Universal Robots URScript: FaiChun_9 Jan_6.script

def Machining1():
  # Default parameters:
  global speed_ms = 0.05
  global speed_rads = 0.75
  global accel_mss = 3
  global accel_radss = 1.2
  global blend_radius_m = 0.0003

  # Add subprograms here
  # Start of main program
  # Program generated by RoboDK v5.6.8 for UR10e on 10/01/2025 10:27:31
  # Using nominal kinematics.
  blend_radius_m = 0.0003
  speed_ms = 0.05
  # set_reference(p[0.325000, -0.070000, 0.000000, 0.000000, 0.000000, 0.000000])
  set_tcp(p[0.000000, 0.000000, 0.252000, 0.000000, 0.000000, 0.000000])
  # Show Tool
  movej([0.540600, -1.409576, -2.440611, -0.862202, 1.570796, 2.111396],accel_radss,speed_rads,0,blend_radius_m)
  movel([0.540600, -1.462244, -2.470081, -0.780064, 1.570796, 2.111396],accel_mss,speed_ms,0,blend_radius_m)
  #SetTool1
  #M_RunCode6
  #SetRPM60000
  speed_ms = 0.05
  #M_RunCode3
  movel([0.540600, -1.485155, -2.481004, -0.746230, 1.570796, 2.111396],accel_mss,speed_ms,0,blend_radius_m)
  speed_ms = 0.003
  movel([0.540600, -1.491068, -2.483663, -0.737658, 1.570796, 2.111396],accel_mss,speed_ms,0,blend_radius_m)
  speed_ms = 0.007
  movel([0.231188, -1.485347, -2.488632, -0.738410, 1.570796, 1.801984],accel_mss,speed_ms,0,blend_radius_m)
  movel([0.347864, -1.099241, -2.719319, -0.893829, 1.570796, 1.918660],accel_mss,speed_ms,0,blend_radius_m)
  movel([0.790744, -1.114546, -2.713470, -0.884373, 1.570796, 2.361541],accel_mss,speed_ms,0,blend_radius_m)
  movel([0.540600, -1.491068, -2.483663, -0.737658, 1.570796, 2.111396],accel_mss,speed_ms,0,blend_radius_m)
  speed_ms = 0.003
  movel([0.540600, -1.485155, -2.481004, -0.746230, 1.570796, 2.111396],accel_mss,speed_ms,0,blend_radius_m)
  speed_ms = 0.05
  movel([0.540600, -1.462244, -2.470081, -0.780064, 1.570796, 2.111396],accel_mss,speed_ms,0,blend_radius_m)
  #M_RunCode9
  movel([0.540492, -1.452284, -2.478323, -0.781782, 1.570796, 2.111289],accel_mss,speed_ms,0,blend_radius_m)
  #M_RunCode3
  movel([0.540492, -1.475406, -2.489363, -0.747620, 1.570796, 2.111289],accel_mss,speed_ms,0,blend_radius_m)
  speed_ms = 0.003
  movel([0.540492, -1.481377, -2.492050, -0.738962, 1.570796, 2.111289],accel_mss,speed_ms,0,blend_radius_m)
  speed_ms = 0.007
  movel([0.536155, -1.480632, -2.492689, -0.739069, 1.570796, 2.106951],accel_mss,speed_ms,0,blend_radius_m)
  movel([0.533586, -1.484990, -2.488940, -0.738459, 1.570796, 2.104382],accel_mss,speed_ms,0,blend_radius_m)
  movel([0.527159, -1.483935, -2.489850, -0.738604, 1.570796, 2.097955],accel_mss,speed_ms,0,blend_radius_m)
  movel([0.529703, -1.479563, -2.493604, -0.739223, 1.570796, 2.100499],accel_mss,speed_ms,0,blend_radius_m)
  movel([0.527435, -1.479199, -2.493915, -0.739276, 1.570796, 2.098231],accel_mss,speed_ms,0,blend_radius_m)
  movel([0.524898, -1.483575, -2.490161, -0.738654, 1.570796, 2.095694],accel_mss,speed_ms,0,blend_radius_m)
  movel([0.519478, -1.482738, -2.490881, -0.738770, 1.570796, 2.090274],accel_mss,speed_ms,0,blend_radius_m)
  movel([0.518427, -1.482577, -2.491019, -0.738793, 1.570796, 2.089223],accel_mss,speed_ms,0,blend_radius_m)
  movel([0.522154, -1.476073, -2.496578, -0.739738, 1.570796, 2.092951],accel_mss,speed_ms,0,blend_radius_m)
  movel([0.526552, -1.476753, -2.496000, -0.739636, 1.570796, 2.097348],accel_mss,speed_ms,0,blend_radius_m)
  movel([0.527881, -1.474461, -2.497945, -0.739983, 1.570796, 2.098677],accel_mss,speed_ms,0,blend_radius_m)
  movel([0.521180, -1.473430, -2.498818, -0.740141, 1.570796, 2.091976],accel_mss,speed_ms,0,blend_radius_m)
  movel([0.516149, -1.482240, -2.491309, -0.738840, 1.570796, 2.086946],accel_mss,speed_ms,0,blend_radius_m)
  movel([0.515092, -1.482086, -2.491441, -0.738862, 1.570796, 2.085888],accel_mss,speed_ms,0,blend_radius_m)
  movel([0.392568, -1.472171, -2.499881, -0.740337, 1.570796, 1.963364],accel_mss,speed_ms,0,blend_radius_m)
  movel([0.261942, -1.477589, -2.495288, -0.739512, 1.570796, 1.832738],accel_mss,speed_ms,0,blend_radius_m)
  movel([0.264591, -1.468670, -2.502825, -0.740895, 1.570796, 1.835387],accel_mss,speed_ms,0,blend_radius_m)
  movel([0.257067, -1.469444, -2.502175, -0.740770, 1.570796, 1.827863],accel_mss,speed_ms,0,blend_radius_m)
  movel([0.256391, -1.471766, -2.500222, -0.740401, 1.570796, 1.827188],accel_mss,speed_ms,0,blend_radius_m)
  movel([0.261332, -1.471251, -2.500656, -0.740482, 1.570796, 1.832129],accel_mss,speed_ms,0,blend_radius_m)
  movel([0.259390, -1.477836, -2.495078, -0.739475, 1.570796, 1.830187],accel_mss,speed_ms,0,blend_radius_m)
  movel([0.258210, -1.477956, -2.494975, -0.739458, 1.570796, 1.829007],accel_mss,speed_ms,0,blend_radius_m)
  movel([0.252127, -1.478591, -2.494434, -0.739364, 1.570796, 1.822923],accel_mss,speed_ms,0,blend_radius_m)
  movel([0.253398, -1.474162, -2.498199, -0.740029, 1.570796, 1.824194],accel_mss,speed_ms,0,blend_radius_m)
  movel([0.250836, -1.474438, -2.497965, -0.739986, 1.570796, 1.821633],accel_mss,speed_ms,0,blend_radius_m)
  movel([0.249578, -1.478866, -2.494199, -0.739324, 1.570796, 1.820375],accel_mss,speed_ms,0,blend_radius_m)
  movel([0.242307, -1.479680, -2.493504, -0.739206, 1.570796, 1.813103],accel_mss,speed_ms,0,blend_radius_m)
  movel([0.243527, -1.475262, -2.497266, -0.739861, 1.570796, 1.814323],accel_mss,speed_ms,0,blend_radius_m)
  movel([0.238589, -1.475844, -2.496772, -0.739773, 1.570796, 1.809385],accel_mss,speed_ms,0,blend_radius_m)
  movel([0.240380, -1.469260, -2.502330, -0.740799, 1.570796, 1.811176],accel_mss,speed_ms,0,blend_radius_m)
  movel([0.245358, -1.468668, -2.502826, -0.740895, 1.570796, 1.816154],accel_mss,speed_ms,0,blend_radius_m)
  movel([0.246004, -1.466343, -2.504771, -0.741276, 1.570796, 1.816800],accel_mss,speed_ms,0,blend_radius_m)
  movel([0.241015, -1.466936, -2.504276, -0.741178, 1.570796, 1.811811],accel_mss,speed_ms,0,blend_radius_m)
  movel([0.242546, -1.461356, -2.508913, -0.742121, 1.570796, 1.813342],accel_mss,speed_ms,0,blend_radius_m)
  movel([0.242845, -1.460267, -2.509812, -0.742310, 1.570796, 1.813642],accel_mss,speed_ms,0,blend_radius_m)
  movel([0.250292, -1.459376, -2.510546, -0.742467, 1.570796, 1.821088],accel_mss,speed_ms,0,blend_radius_m)
  movel([0.249014, -1.463897, -2.506806, -0.741685, 1.570796, 1.819810],accel_mss,speed_ms,0,blend_radius_m)
  movel([0.251610, -1.463600, -2.507053, -0.741736, 1.570796, 1.822406],accel_mss,speed_ms,0,blend_radius_m)
  movel([0.253577, -1.456716, -2.512732, -0.742941, 1.570796, 1.824373],accel_mss,speed_ms,0,blend_radius_m)
  movel([0.243495, -1.457910, -2.511752, -0.742727, 1.570796, 1.814291],accel_mss,speed_ms,0,blend_radius_m)
  movel([0.283133, -1.321596, -2.609965, -0.780829, 1.570796, 1.853929],accel_mss,speed_ms,0,blend_radius_m)
  movel([0.338490, -1.148112, -2.699863, -0.864413, 1.570796, 1.909286],accel_mss,speed_ms,0,blend_radius_m)
  movel([0.339093, -1.146307, -2.700623, -0.865459, 1.570796, 1.909889],accel_mss,speed_ms,0,blend_radius_m)
  movel([0.353258, -1.143604, -2.701755, -0.867030, 1.570796, 1.924055],accel_mss,speed_ms,0,blend_radius_m)
  movel([0.357266, -1.132009, -2.706527, -0.873852, 1.570796, 1.928063],accel_mss,speed_ms,0,blend_radius_m)
  movel([0.353555, -1.132710, -2.706243, -0.873436, 1.570796, 1.924351],accel_mss,speed_ms,0,blend_radius_m)
  movel([0.350931, -1.140355, -2.703106, -0.868929, 1.570796, 1.921727],accel_mss,speed_ms,0,blend_radius_m)
  movel([0.340411, -1.142384, -2.702263, -0.867742, 1.570796, 1.911208],accel_mss,speed_ms,0,blend_radius_m)
  movel([0.341015, -1.140566, -2.703018, -0.868805, 1.570796, 1.911811],accel_mss,speed_ms,0,blend_radius_m)
  movel([0.344182, -1.131093, -2.706899, -0.874397, 1.570796, 1.914978],accel_mss,speed_ms,0,blend_radius_m)
  movel([0.351373, -1.129671, -2.707474, -0.875244, 1.570796, 1.922170],accel_mss,speed_ms,0,blend_radius_m)
  movel([0.352747, -1.125647, -2.709091, -0.877652, 1.570796, 1.923543],accel_mss,speed_ms,0,blend_radius_m)
  movel([0.345526, -1.127083, -2.708515, -0.876791, 1.570796, 1.916323],accel_mss,speed_ms,0,blend_radius_m)
  movel([0.349422, -1.115504, -2.713097, -0.883789, 1.570796, 1.920218],accel_mss,speed_ms,0,blend_radius_m)
  movel([0.356727, -1.114025, -2.713673, -0.884691, 1.570796, 1.927524],accel_mss,speed_ms,0,blend_radius_m)
  movel([0.359466, -1.106053, -2.716742, -0.889593, 1.570796, 1.930262],accel_mss,speed_ms,0,blend_radius_m)
  movel([0.370357, -1.103908, -2.717558, -0.890922, 1.570796, 1.941153],accel_mss,speed_ms,0,blend_radius_m)
  movel([0.367527, -1.111926, -2.714487, -0.885976, 1.570796, 1.938324],accel_mss,speed_ms,0,blend_radius_m)
  movel([0.371310, -1.111216, -2.714761, -0.886412, 1.570796, 1.942106],accel_mss,speed_ms,0,blend_radius_m)
  movel([0.374169, -1.103183, -2.717833, -0.891372, 1.570796, 1.944966],accel_mss,speed_ms,0,blend_radius_m)
  movel([0.385027, -1.101192, -2.718585, -0.892612, 1.570796, 1.955823],accel_mss,speed_ms,0,blend_radius_m)
  movel([0.380684, -1.113104, -2.714031, -0.885255, 1.570796, 1.951481],accel_mss,speed_ms,0,blend_radius_m)
  movel([0.373438, -1.114398, -2.713528, -0.884463, 1.570796, 1.944234],accel_mss,speed_ms,0,blend_radius_m)
  movel([0.371969, -1.118508, -2.711920, -0.881961, 1.570796, 1.942765],accel_mss,speed_ms,0,blend_radius_m)
  movel([0.382929, -1.116581, -2.712676, -0.883132, 1.570796, 1.953725],accel_mss,speed_ms,0,blend_radius_m)
  movel([0.388829, -1.100520, -2.718838, -0.893030, 1.570796, 1.959625],accel_mss,speed_ms,0,blend_radius_m)
  movel([0.580174, -1.086020, -2.724199, -0.902169, 1.570796, 2.150970],accel_mss,speed_ms,0,blend_radius_m)
  movel([0.749145, -1.112705, -2.714185, -0.885499, 1.570796, 2.319942],accel_mss,speed_ms,0,blend_radius_m)
  movel([0.738673, -1.128310, -2.708023, -0.876057, 1.570796, 2.309469],accel_mss,speed_ms,0,blend_radius_m)
  movel([0.747236, -1.130824, -2.707008, -0.874557, 1.570796, 2.318032],accel_mss,speed_ms,0,blend_radius_m)
  movel([0.749941, -1.126842, -2.708612, -0.876935, 1.570796, 2.320738],accel_mss,speed_ms,0,blend_radius_m)
  movel([0.744304, -1.125159, -2.709286, -0.877945, 1.570796, 2.315100],accel_mss,speed_ms,0,blend_radius_m)
  movel([0.752109, -1.113600, -2.713838, -0.884951, 1.570796, 2.322905],accel_mss,speed_ms,0,blend_radius_m)
  movel([0.753475, -1.114012, -2.713678, -0.884699, 1.570796, 2.324272],accel_mss,speed_ms,0,blend_radius_m)
  movel([0.760489, -1.116181, -2.712832, -0.883375, 1.570796, 2.331285],accel_mss,speed_ms,0,blend_radius_m)
  movel([0.755172, -1.123962, -2.709763, -0.878664, 1.570796, 2.325968],accel_mss,speed_ms,0,blend_radius_m)
  movel([0.758077, -1.124873, -2.709400, -0.878116, 1.570796, 2.328873],accel_mss,speed_ms,0,blend_radius_m)
  movel([0.763409, -1.117111, -2.712468, -0.882809, 1.570796, 2.334206],accel_mss,speed_ms,0,blend_radius_m)
  movel([0.771667, -1.119832, -2.711399, -0.881158, 1.570796, 2.342463],accel_mss,speed_ms,0,blend_radius_m)
  movel([0.766309, -1.127539, -2.708332, -0.876518, 1.570796, 2.337105],accel_mss,speed_ms,0,blend_radius_m)
  movel([0.771815, -1.129393, -2.707586, -0.875410, 1.570796, 2.342612],accel_mss,speed_ms,0,blend_radius_m)
  movel([0.763990, -1.140583, -2.703011, -0.868795, 1.570796, 2.334786],accel_mss,speed_ms,0,blend_radius_m)
  movel([0.758513, -1.138781, -2.703756, -0.869852, 1.570796, 2.329309],accel_mss,speed_ms,0,blend_radius_m)
  movel([0.755817, -1.142675, -2.702142, -0.867572, 1.570796, 2.326613],accel_mss,speed_ms,0,blend_radius_m)
  movel([0.761284, -1.144460, -2.701397, -0.866532, 1.570796, 2.332081],accel_mss,speed_ms,0,blend_radius_m)
  movel([0.754898, -1.153625, -2.697523, -0.861241, 1.570796, 2.325695],accel_mss,speed_ms,0,blend_radius_m)
  movel([0.753674, -1.155384, -2.696769, -0.860235, 1.570796, 2.324470],accel_mss,speed_ms,0,blend_radius_m)
  movel([0.745605, -1.152827, -2.697863, -0.861698, 1.570796, 2.316402],accel_mss,speed_ms,0,blend_radius_m)
  movel([0.750697, -1.145425, -2.700993, -0.865971, 1.570796, 2.321494],accel_mss,speed_ms,0,blend_radius_m)
  movel([0.747837, -1.144533, -2.701367, -0.866489, 1.570796, 2.318634],accel_mss,speed_ms,0,blend_radius_m)
  movel([0.740145, -1.155770, -2.696604, -0.860015, 1.570796, 2.310941],accel_mss,speed_ms,0,blend_radius_m)
  movel([0.751042, -1.159170, -2.695138, -0.858082, 1.570796, 2.321838],accel_mss,speed_ms,0,blend_radius_m)
  movel([0.635581, -1.329799, -2.604798, -0.777792, 1.570796, 2.206378],accel_mss,speed_ms,0,blend_radius_m)
  movel([0.551105, -1.463690, -2.506978, -0.741720, 1.570796, 2.121901],accel_mss,speed_ms,0,blend_radius_m)
  movel([0.542267, -1.462159, -2.508248, -0.741982, 1.570796, 2.113063],accel_mss,speed_ms,0,blend_radius_m)
  movel([0.538244, -1.468952, -2.502588, -0.740849, 1.570796, 2.109040],accel_mss,speed_ms,0,blend_radius_m)
  movel([0.540528, -1.469337, -2.502265, -0.740787, 1.570796, 2.111324],accel_mss,speed_ms,0,blend_radius_m)
  movel([0.543178, -1.464878, -2.505991, -0.741520, 1.570796, 2.113974],accel_mss,speed_ms,0,blend_radius_m)
  movel([0.549694, -1.466015, -2.505044, -0.741330, 1.570796, 2.120491],accel_mss,speed_ms,0,blend_radius_m)
  movel([0.549048, -1.467088, -2.504148, -0.741153, 1.570796, 2.119844],accel_mss,speed_ms,0,blend_radius_m)
  movel([0.545741, -1.472593, -2.499525, -0.740271, 1.570796, 2.116537],accel_mss,speed_ms,0,blend_radius_m)
  movel([0.541370, -1.471831, -2.500168, -0.740390, 1.570796, 2.112167],accel_mss,speed_ms,0,blend_radius_m)
  movel([0.540008, -1.474125, -2.498230, -0.740034, 1.570796, 2.110804],accel_mss,speed_ms,0,blend_radius_m)
  movel([0.544370, -1.474884, -2.497587, -0.739918, 1.570796, 2.115167],accel_mss,speed_ms,0,blend_radius_m)
  movel([0.540492, -1.481377, -2.492050, -0.738962, 1.570796, 2.111289],accel_mss,speed_ms,0,blend_radius_m)
  speed_ms = 0.003
  movel([0.540492, -1.475406, -2.489363, -0.747620, 1.570796, 2.111289],accel_mss,speed_ms,0,blend_radius_m)
  speed_ms = 0.05
  movel([0.540492, -1.452284, -2.478323, -0.781782, 1.570796, 2.111289],accel_mss,speed_ms,0,blend_radius_m)
  #M_RunCode9
  movel([0.384099, -1.143946, -2.667631, -0.900812, 1.570796, 1.954895],accel_mss,speed_ms,0,blend_radius_m)
  #M_RunCode3
  movel([0.384099, -1.171719, -2.682638, -0.858032, 1.570796, 1.954895],accel_mss,speed_ms,0,blend_radius_m)
  speed_ms = 0.003
  movel([0.384099, -1.179045, -2.686328, -0.847016, 1.570796, 1.954895],accel_mss,speed_ms,0,blend_radius_m)
  speed_ms = 0.007
  movel([0.371180, -1.190123, -2.681237, -0.841029, 1.570796, 1.941977],accel_mss,speed_ms,0,blend_radius_m)
  movel([0.353670, -1.164627, -2.692759, -0.855002, 1.570796, 1.924466],accel_mss,speed_ms,0,blend_radius_m)
  movel([0.354978, -1.163450, -2.693275, -0.855664, 1.570796, 1.925774],accel_mss,speed_ms,0,blend_radius_m)
  movel([0.358519, -1.160754, -2.694450, -0.857185, 1.570796, 1.929315],accel_mss,speed_ms,0,blend_radius_m)
  movel([0.362422, -1.158698, -2.695342, -0.858349, 1.570796, 1.933218],accel_mss,speed_ms,0,blend_radius_m)
  movel([0.366466, -1.157207, -2.695985, -0.859196, 1.570796, 1.937262],accel_mss,speed_ms,0,blend_radius_m)
  movel([0.370429, -1.156192, -2.696422, -0.859774, 1.570796, 1.941225],accel_mss,speed_ms,0,blend_radius_m)
  movel([0.380760, -1.154569, -2.697119, -0.860701, 1.570796, 1.951557],accel_mss,speed_ms,0,blend_radius_m)
  movel([0.390288, -1.153250, -2.697683, -0.861456, 1.570796, 1.961084],accel_mss,speed_ms,0,blend_radius_m)
  movel([0.393974, -1.152407, -2.698042, -0.861939, 1.570796, 1.964770],accel_mss,speed_ms,0,blend_radius_m)
  movel([0.397663, -1.151161, -2.698572, -0.862655, 1.570796, 1.968460],accel_mss,speed_ms,0,blend_radius_m)
  movel([0.401177, -1.149434, -2.699305, -0.863650, 1.570796, 1.971974],accel_mss,speed_ms,0,blend_radius_m)
  movel([0.404336, -1.147153, -2.700267, -0.864968, 1.570796, 1.975133],accel_mss,speed_ms,0,blend_radius_m)
  movel([0.407651, -1.143740, -2.701698, -0.866951, 1.570796, 1.978447],accel_mss,speed_ms,0,blend_radius_m)
  movel([0.408788, -1.142051, -2.702402, -0.867936, 1.570796, 1.979584],accel_mss,speed_ms,0,blend_radius_m)
  movel([0.409576, -1.140378, -2.703096, -0.868915, 1.570796, 1.980372],accel_mss,speed_ms,0,blend_radius_m)
  movel([0.410196, -1.137359, -2.704342, -0.870688, 1.570796, 1.980993],accel_mss,speed_ms,0,blend_radius_m)
  movel([0.409610, -1.134976, -2.705319, -0.872094, 1.570796, 1.980407],accel_mss,speed_ms,0,blend_radius_m)
  movel([0.408647, -1.133848, -2.705779, -0.872762, 1.570796, 1.979444],accel_mss,speed_ms,0,blend_radius_m)
  movel([0.407469, -1.133422, -2.705953, -0.873014, 1.570796, 1.978266],accel_mss,speed_ms,0,blend_radius_m)
  movel([0.406201, -1.133623, -2.705871, -0.872895, 1.570796, 1.976997],accel_mss,speed_ms,0,blend_radius_m)
  movel([0.404968, -1.134393, -2.705557, -0.872439, 1.570796, 1.975765],accel_mss,speed_ms,0,blend_radius_m)
  movel([0.403605, -1.136287, -2.704782, -0.871320, 1.570796, 1.974401],accel_mss,speed_ms,0,blend_radius_m)
  movel([0.402385, -1.138186, -2.704001, -0.870202, 1.570796, 1.973181],accel_mss,speed_ms,0,blend_radius_m)
  movel([0.400444, -1.140181, -2.703178, -0.869031, 1.570796, 1.971241],accel_mss,speed_ms,0,blend_radius_m)
  movel([0.397817, -1.141968, -2.702436, -0.867985, 1.570796, 1.968613],accel_mss,speed_ms,0,blend_radius_m)
  movel([0.395422, -1.142572, -2.702185, -0.867632, 1.570796, 1.966218],accel_mss,speed_ms,0,blend_radius_m)
  movel([0.393436, -1.142139, -2.702365, -0.867885, 1.570796, 1.964232],accel_mss,speed_ms,0,blend_radius_m)
  movel([0.392041, -1.140812, -2.702916, -0.868661, 1.570796, 1.962837],accel_mss,speed_ms,0,blend_radius_m)
  movel([0.391392, -1.138828, -2.703737, -0.869824, 1.570796, 1.962188],accel_mss,speed_ms,0,blend_radius_m)
  movel([0.391640, -1.136425, -2.704725, -0.871238, 1.570796, 1.962436],accel_mss,speed_ms,0,blend_radius_m)
  movel([0.392852, -1.133853, -2.705777, -0.872758, 1.570796, 1.963649],accel_mss,speed_ms,0,blend_radius_m)
  movel([0.395102, -1.131371, -2.706786, -0.874232, 1.570796, 1.965898],accel_mss,speed_ms,0,blend_radius_m)
  movel([0.397379, -1.129656, -2.707480, -0.875253, 1.570796, 1.968175],accel_mss,speed_ms,0,blend_radius_m)
  movel([0.399624, -1.128553, -2.707925, -0.875911, 1.570796, 1.970420],accel_mss,speed_ms,0,blend_radius_m)
  movel([0.401834, -1.128068, -2.708120, -0.876202, 1.570796, 1.972630],accel_mss,speed_ms,0,blend_radius_m)
  movel([0.404002, -1.128203, -2.708066, -0.876121, 1.570796, 1.974798],accel_mss,speed_ms,0,blend_radius_m)
  movel([0.406053, -1.128886, -2.707791, -0.875713, 1.570796, 1.976850],accel_mss,speed_ms,0,blend_radius_m)
  movel([0.407900, -1.130046, -2.707322, -0.875020, 1.570796, 1.978697],accel_mss,speed_ms,0,blend_radius_m)
  movel([0.410999, -1.133777, -2.705808, -0.872804, 1.570796, 1.981795],accel_mss,speed_ms,0,blend_radius_m)
  movel([0.412374, -1.136716, -2.704606, -0.871067, 1.570796, 1.983170],accel_mss,speed_ms,0,blend_radius_m)
  movel([0.413232, -1.139861, -2.703310, -0.869218, 1.570796, 1.984028],accel_mss,speed_ms,0,blend_radius_m)
  movel([0.413580, -1.143201, -2.701923, -0.867265, 1.570796, 1.984376],accel_mss,speed_ms,0,blend_radius_m)
  movel([0.413422, -1.146734, -2.700444, -0.865211, 1.570796, 1.984218],accel_mss,speed_ms,0,blend_radius_m)
  movel([0.412572, -1.150319, -2.698930, -0.863140, 1.570796, 1.983368],accel_mss,speed_ms,0,blend_radius_m)
  movel([0.410842, -1.153822, -2.697438, -0.861128, 1.570796, 1.981638],accel_mss,speed_ms,0,blend_radius_m)
  movel([0.408237, -1.157248, -2.695968, -0.859173, 1.570796, 1.979033],accel_mss,speed_ms,0,blend_radius_m)
  movel([0.404766, -1.160594, -2.694520, -0.857275, 1.570796, 1.975563],accel_mss,speed_ms,0,blend_radius_m)
  movel([0.401302, -1.163173, -2.693396, -0.855820, 1.570796, 1.972098],accel_mss,speed_ms,0,blend_radius_m)
  movel([0.397796, -1.165070, -2.692565, -0.854754, 1.570796, 1.968592],accel_mss,speed_ms,0,blend_radius_m)
  movel([0.394330, -1.166408, -2.691977, -0.854005, 1.570796, 1.965126],accel_mss,speed_ms,0,blend_radius_m)
  movel([0.391000, -1.167299, -2.691584, -0.853506, 1.570796, 1.961796],accel_mss,speed_ms,0,blend_radius_m)
  movel([0.383085, -1.168489, -2.691058, -0.852842, 1.570796, 1.953882],accel_mss,speed_ms,0,blend_radius_m)
  movel([0.375587, -1.169704, -2.690520, -0.852166, 1.570796, 1.946383],accel_mss,speed_ms,0,blend_radius_m)
  movel([0.372556, -1.170542, -2.690147, -0.851700, 1.570796, 1.943353],accel_mss,speed_ms,0,blend_radius_m)
  movel([0.369459, -1.171768, -2.689601, -0.851020, 1.570796, 1.940255],accel_mss,speed_ms,0,blend_radius_m)
  movel([0.366399, -1.173459, -2.688845, -0.850085, 1.570796, 1.937196],accel_mss,speed_ms,0,blend_radius_m)
  movel([0.363487, -1.175689, -2.687844, -0.848856, 1.570796, 1.934283],accel_mss,speed_ms,0,blend_radius_m)
  movel([0.364141, -1.176646, -2.687413, -0.848330, 1.570796, 1.934937],accel_mss,speed_ms,0,blend_radius_m)
  movel([0.366146, -1.179126, -2.686291, -0.846972, 1.570796, 1.936943],accel_mss,speed_ms,0,blend_radius_m)
  movel([0.368319, -1.180933, -2.685469, -0.845986, 1.570796, 1.939115],accel_mss,speed_ms,0,blend_radius_m)
  movel([0.370657, -1.182078, -2.684947, -0.845364, 1.570796, 1.941454],accel_mss,speed_ms,0,blend_radius_m)
  movel([0.373172, -1.182554, -2.684729, -0.845105, 1.570796, 1.943968],accel_mss,speed_ms,0,blend_radius_m)
  movel([0.375804, -1.182447, -2.684778, -0.845164, 1.570796, 1.946600],accel_mss,speed_ms,0,blend_radius_m)
  movel([0.378498, -1.181829, -2.685061, -0.845499, 1.570796, 1.949294],accel_mss,speed_ms,0,blend_radius_m)
  movel([0.381261, -1.180696, -2.685577, -0.846115, 1.570796, 1.952058],accel_mss,speed_ms,0,blend_radius_m)
  movel([0.384099, -1.179045, -2.686328, -0.847016, 1.570796, 1.954895],accel_mss,speed_ms,0,blend_radius_m)
  speed_ms = 0.003
  movel([0.384099, -1.171719, -2.682638, -0.858032, 1.570796, 1.954895],accel_mss,speed_ms,0,blend_radius_m)
  speed_ms = 0.05
  movel([0.384099, -1.143946, -2.667631, -0.900812, 1.570796, 1.954895],accel_mss,speed_ms,0,blend_radius_m)
  #M_RunCode9
  movel([0.391981, -1.155983, -2.662339, -0.894068, 1.570796, 1.962777],accel_mss,speed_ms,0,blend_radius_m)
  #M_RunCode3
  movel([0.391981, -1.183682, -2.677188, -0.851519, 1.570796, 1.962777],accel_mss,speed_ms,0,blend_radius_m)
  speed_ms = 0.003
  movel([0.391981, -1.190981, -2.680837, -0.840571, 1.570796, 1.962777],accel_mss,speed_ms,0,blend_radius_m)
  speed_ms = 0.007
  movel([0.401981, -1.182312, -2.684840, -0.845237, 1.570796, 1.972777],accel_mss,speed_ms,0,blend_radius_m)
  movel([0.412364, -1.173981, -2.688611, -0.849796, 1.570796, 1.983160],accel_mss,speed_ms,0,blend_radius_m)
  movel([0.420048, -1.168557, -2.691028, -0.852804, 1.570796, 1.990844],accel_mss,speed_ms,0,blend_radius_m)
  movel([0.422893, -1.166993, -2.691719, -0.853677, 1.570796, 1.993689],accel_mss,speed_ms,0,blend_radius_m)
  movel([0.425127, -1.166238, -2.692052, -0.854100, 1.570796, 1.995924],accel_mss,speed_ms,0,blend_radius_m)
  movel([0.426748, -1.166298, -2.692025, -0.854066, 1.570796, 1.997544],accel_mss,speed_ms,0,blend_radius_m)
  movel([0.427747, -1.167174, -2.691639, -0.853576, 1.570796, 1.998543],accel_mss,speed_ms,0,blend_radius_m)
  movel([0.428014, -1.168646, -2.690988, -0.852754, 1.570796, 1.998811],accel_mss,speed_ms,0,blend_radius_m)
  movel([0.427442, -1.170502, -2.690165, -0.851722, 1.570796, 1.998239],accel_mss,speed_ms,0,blend_radius_m)
  movel([0.426031, -1.172734, -2.689170, -0.850485, 1.570796, 1.996828],accel_mss,speed_ms,0,blend_radius_m)
  movel([0.423792, -1.175342, -2.688001, -0.849047, 1.570796, 1.994589],accel_mss,speed_ms,0,blend_radius_m)
  movel([0.416876, -1.181935, -2.685012, -0.845442, 1.570796, 1.987672],accel_mss,speed_ms,0,blend_radius_m)
  movel([0.406811, -1.190510, -2.681057, -0.840823, 1.570796, 1.977607],accel_mss,speed_ms,0,blend_radius_m)
  movel([0.396637, -1.198599, -2.677252, -0.836537, 1.570796, 1.967434],accel_mss,speed_ms,0,blend_radius_m)
  movel([0.389261, -1.203802, -2.674767, -0.833820, 1.570796, 1.960057],accel_mss,speed_ms,0,blend_radius_m)
  movel([0.386540, -1.205311, -2.674041, -0.833037, 1.570796, 1.957337],accel_mss,speed_ms,0,blend_radius_m)
  movel([0.384392, -1.206055, -2.673682, -0.832652, 1.570796, 1.955188],accel_mss,speed_ms,0,blend_radius_m)
  movel([0.382806, -1.206040, -2.673689, -0.832660, 1.570796, 1.953602],accel_mss,speed_ms,0,blend_radius_m)
  movel([0.381784, -1.205259, -2.674066, -0.833064, 1.570796, 1.952580],accel_mss,speed_ms,0,blend_radius_m)
  movel([0.381444, -1.203906, -2.674717, -0.833765, 1.570796, 1.952240],accel_mss,speed_ms,0,blend_radius_m)
  movel([0.381917, -1.202164, -2.675553, -0.834672, 1.570796, 1.952713],accel_mss,speed_ms,0,blend_radius_m)
  movel([0.383201, -1.200030, -2.676572, -0.835787, 1.570796, 1.953998],accel_mss,speed_ms,0,blend_radius_m)
  movel([0.385310, -1.197499, -2.677774, -0.837116, 1.570796, 1.956107],accel_mss,speed_ms,0,blend_radius_m)
  movel([0.391981, -1.190981, -2.680837, -0.840571, 1.570796, 1.962777],accel_mss,speed_ms,0,blend_radius_m)
  speed_ms = 0.003
  movel([0.391981, -1.183682, -2.677188, -0.851519, 1.570796, 1.962777],accel_mss,speed_ms,0,blend_radius_m)
  speed_ms = 0.05
  movel([0.391981, -1.155983, -2.662339, -0.894068, 1.570796, 1.962777],accel_mss,speed_ms,0,blend_radius_m)
  #M_RunCode9
  movel([0.382534, -1.154364, -2.663059, -0.894966, 1.570796, 1.953331],accel_mss,speed_ms,0,blend_radius_m)
  #M_RunCode3
  movel([0.382534, -1.182074, -2.677929, -0.852386, 1.570796, 1.953331],accel_mss,speed_ms,0,blend_radius_m)
  speed_ms = 0.003
  movel([0.382534, -1.189377, -2.681584, -0.841428, 1.570796, 1.953331],accel_mss,speed_ms,0,blend_radius_m)
  speed_ms = 0.007
  movel([0.384510, -1.186300, -2.683009, -0.843080, 1.570796, 1.955306],accel_mss,speed_ms,0,blend_radius_m)
  movel([0.386914, -1.183128, -2.684467, -0.844794, 1.570796, 1.957710],accel_mss,speed_ms,0,blend_radius_m)
  movel([0.389736, -1.179922, -2.685929, -0.846537, 1.570796, 1.960532],accel_mss,speed_ms,0,blend_radius_m)
  movel([0.392976, -1.176687, -2.687394, -0.848307, 1.570796, 1.963773],accel_mss,speed_ms,0,blend_radius_m)
  movel([0.396639, -1.173419, -2.688863, -0.850106, 1.570796, 1.967435],accel_mss,speed_ms,0,blend_radius_m)
  movel([0.400453, -1.170358, -2.690229, -0.851802, 1.570796, 1.971250],accel_mss,speed_ms,0,blend_radius_m)
  movel([0.404137, -1.167738, -2.691390, -0.853261, 1.570796, 1.974933],accel_mss,speed_ms,0,blend_radius_m)
  movel([0.407690, -1.165566, -2.692347, -0.854476, 1.570796, 1.978486],accel_mss,speed_ms,0,blend_radius_m)
  movel([0.411102, -1.163850, -2.693100, -0.855439, 1.570796, 1.981898],accel_mss,speed_ms,0,blend_radius_m)
  movel([0.414313, -1.162590, -2.693651, -0.856149, 1.570796, 1.985110],accel_mss,speed_ms,0,blend_radius_m)
  movel([0.417262, -1.161790, -2.694000, -0.856600, 1.570796, 1.988058],accel_mss,speed_ms,0,blend_radius_m)
  movel([0.419951, -1.161449, -2.694148, -0.856792, 1.570796, 1.990747],accel_mss,speed_ms,0,blend_radius_m)
  movel([0.422369, -1.161571, -2.694095, -0.856723, 1.570796, 1.993165],accel_mss,speed_ms,0,blend_radius_m)
  movel([0.424501, -1.162118, -2.693856, -0.856414, 1.570796, 1.995297],accel_mss,speed_ms,0,blend_radius_m)
  movel([0.426315, -1.163065, -2.693443, -0.855881, 1.570796, 1.997111],accel_mss,speed_ms,0,blend_radius_m)
  movel([0.427820, -1.164408, -2.692856, -0.855126, 1.570796, 1.998617],accel_mss,speed_ms,0,blend_radius_m)
  movel([0.429009, -1.166139, -2.692095, -0.854155, 1.570796, 1.999805],accel_mss,speed_ms,0,blend_radius_m)
  movel([0.429838, -1.168160, -2.691203, -0.853025, 1.570796, 2.000634],accel_mss,speed_ms,0,blend_radius_m)
  movel([0.430255, -1.170379, -2.690220, -0.851791, 1.570796, 2.001051],accel_mss,speed_ms,0,blend_radius_m)
  movel([0.430265, -1.172781, -2.689149, -0.850459, 1.570796, 2.001061],accel_mss,speed_ms,0,blend_radius_m)
  movel([0.429867, -1.175374, -2.687986, -0.849029, 1.570796, 2.000663],accel_mss,speed_ms,0,blend_radius_m)
  movel([0.429057, -1.178111, -2.686751, -0.847527, 1.570796, 1.999853],accel_mss,speed_ms,0,blend_radius_m)
  movel([0.427818, -1.180961, -2.685457, -0.845972, 1.570796, 1.998614],accel_mss,speed_ms,0,blend_radius_m)
  movel([0.426158, -1.183915, -2.684106, -0.844368, 1.570796, 1.996955],accel_mss,speed_ms,0,blend_radius_m)
  movel([0.424077, -1.186979, -2.682695, -0.842715, 1.570796, 1.994873],accel_mss,speed_ms,0,blend_radius_m)
  movel([0.421597, -1.190091, -2.681252, -0.841046, 1.570796, 1.992393],accel_mss,speed_ms,0,blend_radius_m)
  movel([0.418745, -1.193188, -2.679805, -0.839396, 1.570796, 1.989541],accel_mss,speed_ms,0,blend_radius_m)
  movel([0.415518, -1.196270, -2.678355, -0.837764, 1.570796, 1.986314],accel_mss,speed_ms,0,blend_radius_m)
  movel([0.411919, -1.199346, -2.676897, -0.836146, 1.570796, 1.982715],accel_mss,speed_ms,0,blend_radius_m)
  movel([0.408214, -1.202196, -2.675537, -0.834655, 1.570796, 1.979010],accel_mss,speed_ms,0,blend_radius_m)
  movel([0.404666, -1.204615, -2.674377, -0.833398, 1.570796, 1.975463],accel_mss,speed_ms,0,blend_radius_m)
  movel([0.401273, -1.206606, -2.673416, -0.832367, 1.570796, 1.972069],accel_mss,speed_ms,0,blend_radius_m)
  movel([0.398024, -1.208172, -2.672657, -0.831560, 1.570796, 1.968821],accel_mss,speed_ms,0,blend_radius_m)
  movel([0.394967, -1.209327, -2.672096, -0.830966, 1.570796, 1.965763],accel_mss,speed_ms,0,blend_radius_m)
  movel([0.392151, -1.210070, -2.671734, -0.830585, 1.570796, 1.962947],accel_mss,speed_ms,0,blend_radius_m)
  movel([0.389569, -1.210403, -2.671572, -0.830414, 1.570796, 1.960365],accel_mss,speed_ms,0,blend_radius_m)
  movel([0.387217, -1.210331, -2.671607, -0.830451, 1.570796, 1.958013],accel_mss,speed_ms,0,blend_radius_m)
  movel([0.385124, -1.209875, -2.671829, -0.830685, 1.570796, 1.955920],accel_mss,speed_ms,0,blend_radius_m)
  movel([0.383309, -1.209055, -2.672228, -0.831106, 1.570796, 1.954105],accel_mss,speed_ms,0,blend_radius_m)
  movel([0.381774, -1.207869, -2.672804, -0.831715, 1.570796, 1.952571],accel_mss,speed_ms,0,blend_radius_m)
  movel([0.380519, -1.206319, -2.673555, -0.832516, 1.570796, 1.951316],accel_mss,speed_ms,0,blend_radius_m)
  movel([0.379600, -1.204481, -2.674441, -0.833467, 1.570796, 1.950397],accel_mss,speed_ms,0,blend_radius_m)
  movel([0.379072, -1.202440, -2.675421, -0.834528, 1.570796, 1.949868],accel_mss,speed_ms,0,blend_radius_m)
  movel([0.378939, -1.200190, -2.676496, -0.835703, 1.570796, 1.949735],accel_mss,speed_ms,0,blend_radius_m)
  movel([0.379206, -1.197729, -2.677665, -0.836995, 1.570796, 1.950002],accel_mss,speed_ms,0,blend_radius_m)
  movel([0.379886, -1.195089, -2.678912, -0.838388, 1.570796, 1.950682],accel_mss,speed_ms,0,blend_radius_m)
  movel([0.380993, -1.192308, -2.680217, -0.839864, 1.570796, 1.951790],accel_mss,speed_ms,0,blend_radius_m)
  movel([0.382534, -1.189377, -2.681584, -0.841428, 1.570796, 1.953331],accel_mss,speed_ms,0,blend_radius_m)
  speed_ms = 0.003
  movel([0.382534, -1.182074, -2.677929, -0.852386, 1.570796, 1.953331],accel_mss,speed_ms,0,blend_radius_m)
  speed_ms = 0.05
  movel([0.382534, -1.154364, -2.663059, -0.894966, 1.570796, 1.953331],accel_mss,speed_ms,0,blend_radius_m)
  #M_RunCode9
  movel([0.494383, -1.389930, -2.526626, -0.795833, 1.570796, 2.065179],accel_mss,speed_ms,0,blend_radius_m)
  #M_RunCode3
  movel([0.494383, -1.414326, -2.538424, -0.759639, 1.570796, 2.065179],accel_mss,speed_ms,0,blend_radius_m)
  speed_ms = 0.003
  movel([0.494383, -1.420647, -2.541300, -0.750441, 1.570796, 2.065179],accel_mss,speed_ms,0,blend_radius_m)
  speed_ms = 0.007
  movel([0.497081, -1.419373, -2.542274, -0.750742, 1.570796, 2.067877],accel_mss,speed_ms,0,blend_radius_m)
  movel([0.499941, -1.418639, -2.542833, -0.750917, 1.570796, 2.070737],accel_mss,speed_ms,0,blend_radius_m)
  movel([0.502829, -1.418338, -2.543062, -0.750988, 1.570796, 2.073625],accel_mss,speed_ms,0,blend_radius_m)
  movel([0.505605, -1.418366, -2.543041, -0.750982, 1.570796, 2.076401],accel_mss,speed_ms,0,blend_radius_m)
  movel([0.512719, -1.419167, -2.542431, -0.750791, 1.570796, 2.083515],accel_mss,speed_ms,0,blend_radius_m)
  movel([0.519252, -1.420019, -2.541780, -0.750589, 1.570796, 2.090049],accel_mss,speed_ms,0,blend_radius_m)
  movel([0.521814, -1.420108, -2.541713, -0.750569, 1.570796, 2.092610],accel_mss,speed_ms,0,blend_radius_m)
  movel([0.524418, -1.419908, -2.541865, -0.750616, 1.570796, 2.095214],accel_mss,speed_ms,0,blend_radius_m)
  movel([0.526952, -1.419333, -2.542304, -0.750752, 1.570796, 2.097748],accel_mss,speed_ms,0,blend_radius_m)
  movel([0.529302, -1.418300, -2.543092, -0.750998, 1.570796, 2.100099],accel_mss,speed_ms,0,blend_radius_m)
  movel([0.531866, -1.416496, -2.544463, -0.751431, 1.570796, 2.102662],accel_mss,speed_ms,0,blend_radius_m)
  movel([0.532796, -1.415514, -2.545207, -0.751668, 1.570796, 2.103592],accel_mss,speed_ms,0,blend_radius_m)
  movel([0.533494, -1.414477, -2.545991, -0.751921, 1.570796, 2.104290],accel_mss,speed_ms,0,blend_radius_m)
  movel([0.534215, -1.412459, -2.547513, -0.752417, 1.570796, 2.105012],accel_mss,speed_ms,0,blend_radius_m)
  movel([0.534067, -1.410667, -2.548859, -0.752863, 1.570796, 2.104864],accel_mss,speed_ms,0,blend_radius_m)
  movel([0.533541, -1.409690, -2.549591, -0.753108, 1.570796, 2.104338],accel_mss,speed_ms,0,blend_radius_m)
  movel([0.532799, -1.409167, -2.549982, -0.753240, 1.570796, 2.103596],accel_mss,speed_ms,0,blend_radius_m)
  movel([0.531934, -1.409071, -2.550054, -0.753264, 1.570796, 2.102730],accel_mss,speed_ms,0,blend_radius_m)
  movel([0.531038, -1.409381, -2.549822, -0.753186, 1.570796, 2.101834],accel_mss,speed_ms,0,blend_radius_m)
  movel([0.529935, -1.410463, -2.549012, -0.752914, 1.570796, 2.100731],accel_mss,speed_ms,0,blend_radius_m)
  movel([0.528924, -1.411578, -2.548175, -0.752636, 1.570796, 2.099720],accel_mss,speed_ms,0,blend_radius_m)
  movel([0.527424, -1.412624, -2.547389, -0.752376, 1.570796, 2.098220],accel_mss,speed_ms,0,blend_radius_m)
  movel([0.525483, -1.413399, -2.546805, -0.752185, 1.570796, 2.096280],accel_mss,speed_ms,0,blend_radius_m)
  movel([0.523822, -1.413373, -2.546824, -0.752192, 1.570796, 2.094618],accel_mss,speed_ms,0,blend_radius_m)
  movel([0.522542, -1.412689, -2.547340, -0.752360, 1.570796, 2.093338],accel_mss,speed_ms,0,blend_radius_m)
  movel([0.521753, -1.411480, -2.548249, -0.752660, 1.570796, 2.092549],accel_mss,speed_ms,0,blend_radius_m)
  movel([0.521531, -1.409947, -2.549399, -0.753043, 1.570796, 2.092327],accel_mss,speed_ms,0,blend_radius_m)
  movel([0.521953, -1.408286, -2.550640, -0.753462, 1.570796, 2.092749],accel_mss,speed_ms,0,blend_radius_m)
  movel([0.523034, -1.406692, -2.551828, -0.753868, 1.570796, 2.093830],accel_mss,speed_ms,0,blend_radius_m)
  movel([0.524792, -1.405362, -2.552817, -0.754210, 1.570796, 2.095589],accel_mss,speed_ms,0,blend_radius_m)
  movel([0.526486, -1.404585, -2.553393, -0.754411, 1.570796, 2.097282],accel_mss,speed_ms,0,blend_radius_m)
  movel([0.528091, -1.404236, -2.553652, -0.754502, 1.570796, 2.098888],accel_mss,speed_ms,0,blend_radius_m)
  movel([0.529608, -1.404316, -2.553592, -0.754481, 1.570796, 2.100405],accel_mss,speed_ms,0,blend_radius_m)
  movel([0.531035, -1.404826, -2.553214, -0.754349, 1.570796, 2.101831],accel_mss,speed_ms,0,blend_radius_m)
  movel([0.532324, -1.405698, -2.552567, -0.754124, 1.570796, 2.103120],accel_mss,speed_ms,0,blend_radius_m)
  movel([0.533433, -1.406868, -2.551698, -0.753824, 1.570796, 2.104229],accel_mss,speed_ms,0,blend_radius_m)
  movel([0.535111, -1.410082, -2.549298, -0.753010, 1.570796, 2.105907],accel_mss,speed_ms,0,blend_radius_m)
  movel([0.535730, -1.412414, -2.547547, -0.752428, 1.570796, 2.106526],accel_mss,speed_ms,0,blend_radius_m)
  movel([0.535987, -1.414790, -2.545754, -0.751845, 1.570796, 2.106783],accel_mss,speed_ms,0,blend_radius_m)
  movel([0.535884, -1.417214, -2.543918, -0.751258, 1.570796, 2.106680],accel_mss,speed_ms,0,blend_radius_m)
  movel([0.535424, -1.419683, -2.542037, -0.750669, 1.570796, 2.106221],accel_mss,speed_ms,0,blend_radius_m)
  movel([0.534495, -1.422065, -2.540215, -0.750110, 1.570796, 2.105292],accel_mss,speed_ms,0,blend_radius_m)
  movel([0.532980, -1.424234, -2.538547, -0.749607, 1.570796, 2.103776],accel_mss,speed_ms,0,blend_radius_m)
  movel([0.530887, -1.426191, -2.537037, -0.749161, 1.570796, 2.101683],accel_mss,speed_ms,0,blend_radius_m)
  movel([0.528209, -1.427943, -2.535681, -0.748765, 1.570796, 2.099005],accel_mss,speed_ms,0,blend_radius_m)
  movel([0.525614, -1.429150, -2.534743, -0.748496, 1.570796, 2.096411],accel_mss,speed_ms,0,blend_radius_m)
  movel([0.523054, -1.429866, -2.534186, -0.748337, 1.570796, 2.093850],accel_mss,speed_ms,0,blend_radius_m)
  movel([0.520575, -1.430192, -2.533932, -0.748265, 1.570796, 2.091372],accel_mss,speed_ms,0,blend_radius_m)
  movel([0.518236, -1.430218, -2.533912, -0.748259, 1.570796, 2.089032],accel_mss,speed_ms,0,blend_radius_m)
  movel([0.512764, -1.429613, -2.534383, -0.748393, 1.570796, 2.083560],accel_mss,speed_ms,0,blend_radius_m)
  movel([0.507570, -1.429093, -2.534787, -0.748508, 1.570796, 2.078366],accel_mss,speed_ms,0,blend_radius_m)
  movel([0.505430, -1.429133, -2.534757, -0.748500, 1.570796, 2.076226],accel_mss,speed_ms,0,blend_radius_m)
  movel([0.503200, -1.429440, -2.534518, -0.748432, 1.570796, 2.073996],accel_mss,speed_ms,0,blend_radius_m)
  movel([0.500938, -1.430091, -2.534011, -0.748287, 1.570796, 2.071735],accel_mss,speed_ms,0,blend_radius_m)
  movel([0.498716, -1.431164, -2.533174, -0.748051, 1.570796, 2.069512],accel_mss,speed_ms,0,blend_radius_m)
  movel([0.499050, -1.431983, -2.532534, -0.747872, 1.570796, 2.069846],accel_mss,speed_ms,0,blend_radius_m)
  movel([0.500128, -1.434162, -2.530827, -0.747400, 1.570796, 2.070924],accel_mss,speed_ms,0,blend_radius_m)
  movel([0.501395, -1.435883, -2.529473, -0.747032, 1.570796, 2.072191],accel_mss,speed_ms,0,blend_radius_m)
  movel([0.502857, -1.437147, -2.528476, -0.746765, 1.570796, 2.073653],accel_mss,speed_ms,0,blend_radius_m)
  movel([0.504510, -1.437959, -2.527835, -0.746595, 1.570796, 2.075306],accel_mss,speed_ms,0,blend_radius_m)
  movel([0.506311, -1.438363, -2.527515, -0.746511, 1.570796, 2.077107],accel_mss,speed_ms,0,blend_radius_m)
  movel([0.508208, -1.438409, -2.527479, -0.746501, 1.570796, 2.079004],accel_mss,speed_ms,0,blend_radius_m)
  movel([0.510207, -1.438094, -2.527728, -0.746567, 1.570796, 2.081003],accel_mss,speed_ms,0,blend_radius_m)
  movel([0.512309, -1.437419, -2.528261, -0.746708, 1.570796, 2.083106],accel_mss,speed_ms,0,blend_radius_m)
  movel([0.502315, -1.443102, -2.523747, -0.745540, 1.570796, 2.073111],accel_mss,speed_ms,0,blend_radius_m)
  movel([0.493365, -1.421248, -2.540841, -0.750300, 1.570796, 2.064162],accel_mss,speed_ms,0,blend_radius_m)
  movel([0.494383, -1.420647, -2.541300, -0.750441, 1.570796, 2.065179],accel_mss,speed_ms,0,blend_radius_m)
  speed_ms = 0.003
  movel([0.494383, -1.414326, -2.538424, -0.759639, 1.570796, 2.065179],accel_mss,speed_ms,0,blend_radius_m)
  speed_ms = 0.05
  movel([0.494383, -1.389930, -2.526626, -0.795833, 1.570796, 2.065179],accel_mss,speed_ms,0,blend_radius_m)
  #M_RunCode9
  movel([0.509612, -1.412120, -2.510078, -0.790191, 1.570796, 2.080409],accel_mss,speed_ms,0,blend_radius_m)
  #M_RunCode3
  movel([0.509612, -1.436073, -2.521602, -0.754714, 1.570796, 2.080409],accel_mss,speed_ms,0,blend_radius_m)
  speed_ms = 0.003
  movel([0.509612, -1.442272, -2.524410, -0.745707, 1.570796, 2.080409],accel_mss,speed_ms,0,blend_radius_m)
  speed_ms = 0.007
  movel([0.511490, -1.441522, -2.525007, -0.745860, 1.570796, 2.082287],accel_mss,speed_ms,0,blend_radius_m)
  movel([0.513128, -1.441532, -2.525000, -0.745858, 1.570796, 2.083924],accel_mss,speed_ms,0,blend_radius_m)
  movel([0.514398, -1.442178, -2.524485, -0.745726, 1.570796, 2.085195],accel_mss,speed_ms,0,blend_radius_m)
  movel([0.515181, -1.443333, -2.523562, -0.745493, 1.570796, 2.085977],accel_mss,speed_ms,0,blend_radius_m)
  movel([0.515399, -1.444801, -2.522388, -0.745200, 1.570796, 2.086195],accel_mss,speed_ms,0,blend_radius_m)
  movel([0.514982, -1.446386, -2.521116, -0.744887, 1.570796, 2.085779],accel_mss,speed_ms,0,blend_radius_m)
  movel([0.513938, -1.447896, -2.519900, -0.744592, 1.570796, 2.084734],accel_mss,speed_ms,0,blend_radius_m)
  movel([0.512272, -1.449136, -2.518900, -0.744353, 1.570796, 2.083068],accel_mss,speed_ms,0,blend_radius_m)
  movel([0.510726, -1.449811, -2.518354, -0.744224, 1.570796, 2.081522],accel_mss,speed_ms,0,blend_radius_m)
  movel([0.509449, -1.450009, -2.518194, -0.744186, 1.570796, 2.080246],accel_mss,speed_ms,0,blend_radius_m)
  movel([0.508135, -1.450311, -2.517949, -0.744128, 1.570796, 2.078931],accel_mss,speed_ms,0,blend_radius_m)
  movel([0.507400, -1.450916, -2.517460, -0.744014, 1.570796, 2.078197],accel_mss,speed_ms,0,blend_radius_m)
  movel([0.506930, -1.451756, -2.516778, -0.743855, 1.570796, 2.077727],accel_mss,speed_ms,0,blend_radius_m)
  movel([0.506762, -1.452683, -2.516025, -0.743681, 1.570796, 2.077558],accel_mss,speed_ms,0,blend_radius_m)
  movel([0.506927, -1.453558, -2.515312, -0.743519, 1.570796, 2.077723],accel_mss,speed_ms,0,blend_radius_m)
  movel([0.507485, -1.454522, -2.514526, -0.743341, 1.570796, 2.078282],accel_mss,speed_ms,0,blend_radius_m)
  movel([0.508303, -1.455228, -2.513950, -0.743211, 1.570796, 2.079099],accel_mss,speed_ms,0,blend_radius_m)
  movel([0.509379, -1.455675, -2.513584, -0.743130, 1.570796, 2.080176],accel_mss,speed_ms,0,blend_radius_m)
  movel([0.510712, -1.455870, -2.513425, -0.743094, 1.570796, 2.081508],accel_mss,speed_ms,0,blend_radius_m)
  movel([0.512224, -1.455797, -2.513485, -0.743108, 1.570796, 2.083021],accel_mss,speed_ms,0,blend_radius_m)
  movel([0.513839, -1.455450, -2.513768, -0.743171, 1.570796, 2.084635],accel_mss,speed_ms,0,blend_radius_m)
  movel([0.515560, -1.454826, -2.514278, -0.743285, 1.570796, 2.086356],accel_mss,speed_ms,0,blend_radius_m)
  movel([0.517386, -1.453926, -2.515013, -0.743451, 1.570796, 2.088182],accel_mss,speed_ms,0,blend_radius_m)
  movel([0.520257, -1.451945, -2.516624, -0.743819, 1.570796, 2.091053],accel_mss,speed_ms,0,blend_radius_m)
  movel([0.522585, -1.449475, -2.518626, -0.744288, 1.570796, 2.093382],accel_mss,speed_ms,0,blend_radius_m)
  movel([0.523520, -1.448065, -2.519765, -0.744560, 1.570796, 2.094316],accel_mss,speed_ms,0,blend_radius_m)
  movel([0.524260, -1.446552, -2.520982, -0.744854, 1.570796, 2.095056],accel_mss,speed_ms,0,blend_radius_m)
  movel([0.525158, -1.443210, -2.523661, -0.745518, 1.570796, 2.095955],accel_mss,speed_ms,0,blend_radius_m)
  movel([0.525179, -1.439539, -2.526583, -0.746267, 1.570796, 2.095975],accel_mss,speed_ms,0,blend_radius_m)
  movel([0.524211, -1.435637, -2.529668, -0.747085, 1.570796, 2.095007],accel_mss,speed_ms,0,blend_radius_m)
  movel([0.539789, -1.427052, -2.536371, -0.748966, 1.570796, 2.110585],accel_mss,speed_ms,0,blend_radius_m)
  movel([0.545461, -1.443958, -2.523063, -0.745368, 1.570796, 2.116257],accel_mss,speed_ms,0,blend_radius_m)
  movel([0.535452, -1.449327, -2.518746, -0.744316, 1.570796, 2.106249],accel_mss,speed_ms,0,blend_radius_m)
  movel([0.537620, -1.447411, -2.520291, -0.744687, 1.570796, 2.108416],accel_mss,speed_ms,0,blend_radius_m)
  movel([0.539396, -1.445076, -2.522167, -0.745145, 1.570796, 2.110192],accel_mss,speed_ms,0,blend_radius_m)
  movel([0.540687, -1.442436, -2.524279, -0.745674, 1.570796, 2.111484],accel_mss,speed_ms,0,blend_radius_m)
  movel([0.541406, -1.439606, -2.526530, -0.746253, 1.570796, 2.112203],accel_mss,speed_ms,0,blend_radius_m)
  movel([0.541489, -1.436695, -2.528833, -0.746861, 1.570796, 2.112285],accel_mss,speed_ms,0,blend_radius_m)
  movel([0.540874, -1.433817, -2.531098, -0.747474, 1.570796, 2.111670],accel_mss,speed_ms,0,blend_radius_m)
  movel([0.529435, -1.440058, -2.526171, -0.746160, 1.570796, 2.100232],accel_mss,speed_ms,0,blend_radius_m)
  movel([0.530293, -1.443522, -2.523411, -0.745455, 1.570796, 2.101089],accel_mss,speed_ms,0,blend_radius_m)
  movel([0.530471, -1.447177, -2.520480, -0.744732, 1.570796, 2.101268],accel_mss,speed_ms,0,blend_radius_m)
  movel([0.529866, -1.450823, -2.517535, -0.744031, 1.570796, 2.100662],accel_mss,speed_ms,0,blend_radius_m)
  movel([0.529229, -1.452573, -2.516114, -0.743702, 1.570796, 2.100025],accel_mss,speed_ms,0,blend_radius_m)
  movel([0.528372, -1.454274, -2.514729, -0.743386, 1.570796, 2.099168],accel_mss,speed_ms,0,blend_radius_m)
  movel([0.527276, -1.455875, -2.513420, -0.743093, 1.570796, 2.098072],accel_mss,speed_ms,0,blend_radius_m)
  movel([0.525923, -1.457328, -2.512230, -0.742831, 1.570796, 2.096719],accel_mss,speed_ms,0,blend_radius_m)
  movel([0.524317, -1.458631, -2.511159, -0.742598, 1.570796, 2.095113],accel_mss,speed_ms,0,blend_radius_m)
  movel([0.522454, -1.459792, -2.510204, -0.742393, 1.570796, 2.093250],accel_mss,speed_ms,0,blend_radius_m)
  movel([0.520506, -1.460724, -2.509434, -0.742230, 1.570796, 2.091302],accel_mss,speed_ms,0,blend_radius_m)
  movel([0.518643, -1.461347, -2.508920, -0.742122, 1.570796, 2.089440],accel_mss,speed_ms,0,blend_radius_m)
  movel([0.516862, -1.461661, -2.508660, -0.742068, 1.570796, 2.087658],accel_mss,speed_ms,0,blend_radius_m)
  movel([0.515163, -1.461668, -2.508654, -0.742067, 1.570796, 2.085960],accel_mss,speed_ms,0,blend_radius_m)
  movel([0.512100, -1.460952, -2.509246, -0.742191, 1.570796, 2.082897],accel_mss,speed_ms,0,blend_radius_m)
  movel([0.509548, -1.459390, -2.510535, -0.742464, 1.570796, 2.080345],accel_mss,speed_ms,0,blend_radius_m)
  movel([0.507542, -1.457189, -2.512344, -0.742856, 1.570796, 2.078338],accel_mss,speed_ms,0,blend_radius_m)
  movel([0.506120, -1.454557, -2.514498, -0.743334, 1.570796, 2.076917],accel_mss,speed_ms,0,blend_radius_m)
  movel([0.505558, -1.452516, -2.516160, -0.743713, 1.570796, 2.076354],accel_mss,speed_ms,0,blend_radius_m)
  movel([0.505383, -1.450221, -2.518022, -0.744145, 1.570796, 2.076179],accel_mss,speed_ms,0,blend_radius_m)
  movel([0.505659, -1.447865, -2.519926, -0.744598, 1.570796, 2.076455],accel_mss,speed_ms,0,blend_radius_m)
  movel([0.506446, -1.445637, -2.521718, -0.745034, 1.570796, 2.077243],accel_mss,speed_ms,0,blend_radius_m)
  movel([0.507761, -1.443713, -2.523259, -0.745417, 1.570796, 2.078557],accel_mss,speed_ms,0,blend_radius_m)
  movel([0.509612, -1.442272, -2.524410, -0.745707, 1.570796, 2.080409],accel_mss,speed_ms,0,blend_radius_m)
  speed_ms = 0.003
  movel([0.509612, -1.436073, -2.521602, -0.754714, 1.570796, 2.080409],accel_mss,speed_ms,0,blend_radius_m)
  speed_ms = 0.05
  movel([0.509612, -1.412120, -2.510078, -0.790191, 1.570796, 2.080409],accel_mss,speed_ms,0,blend_radius_m)
  #M_RunCode9
  movel([0.517025, -1.320922, -2.573739, -0.817728, 1.570796, 2.087821],accel_mss,speed_ms,0,blend_radius_m)
  #M_RunCode3
  movel([0.517025, -1.346591, -2.586414, -0.779384, 1.570796, 2.087821],accel_mss,speed_ms,0,blend_radius_m)
  speed_ms = 0.003
  movel([0.517025, -1.353271, -2.589511, -0.769607, 1.570796, 2.087821],accel_mss,speed_ms,0,blend_radius_m)
  speed_ms = 0.007
  movel([0.513857, -1.353859, -2.589119, -0.769412, 1.570796, 2.084654],accel_mss,speed_ms,0,blend_radius_m)
  movel([0.510784, -1.353806, -2.589154, -0.769429, 1.570796, 2.081580],accel_mss,speed_ms,0,blend_radius_m)
  movel([0.507871, -1.353220, -2.589545, -0.769624, 1.570796, 2.078668],accel_mss,speed_ms,0,blend_radius_m)
  movel([0.505181, -1.352209, -2.590219, -0.769961, 1.570796, 2.075978],accel_mss,speed_ms,0,blend_radius_m)
  movel([0.502784, -1.350876, -2.591105, -0.770407, 1.570796, 2.073580],accel_mss,speed_ms,0,blend_radius_m)
  movel([0.504597, -1.347224, -2.593522, -0.771643, 1.570796, 2.075394],accel_mss,speed_ms,0,blend_radius_m)
  movel([0.507463, -1.343318, -2.596086, -0.772985, 1.570796, 2.078259],accel_mss,speed_ms,0,blend_radius_m)
  movel([0.511084, -1.339508, -2.598566, -0.774315, 1.570796, 2.081881],accel_mss,speed_ms,0,blend_radius_m)
  movel([0.515153, -1.336160, -2.600729, -0.775499, 1.570796, 2.085949],accel_mss,speed_ms,0,blend_radius_m)
  movel([0.519346, -1.333645, -2.602345, -0.776399, 1.570796, 2.090142],accel_mss,speed_ms,0,blend_radius_m)
  movel([0.521387, -1.332816, -2.602876, -0.776698, 1.570796, 2.092183],accel_mss,speed_ms,0,blend_radius_m)
  movel([0.523335, -1.332335, -2.603183, -0.776871, 1.570796, 2.094131],accel_mss,speed_ms,0,blend_radius_m)
  movel([0.525151, -1.332246, -2.603239, -0.776903, 1.570796, 2.095947],accel_mss,speed_ms,0,blend_radius_m)
  movel([0.526785, -1.332598, -2.603015, -0.776776, 1.570796, 2.097581],accel_mss,speed_ms,0,blend_radius_m)
  movel([0.528204, -1.333429, -2.602483, -0.776477, 1.570796, 2.099000],accel_mss,speed_ms,0,blend_radius_m)
  movel([0.529362, -1.334787, -2.601613, -0.775989, 1.570796, 2.100158],accel_mss,speed_ms,0,blend_radius_m)
  movel([0.530223, -1.337369, -2.599950, -0.775070, 1.570796, 2.101019],accel_mss,speed_ms,0,blend_radius_m)
  movel([0.529939, -1.340263, -2.598076, -0.774050, 1.570796, 2.100735],accel_mss,speed_ms,0,blend_radius_m)
  movel([0.528649, -1.343348, -2.596066, -0.772975, 1.570796, 2.099445],accel_mss,speed_ms,0,blend_radius_m)
  movel([0.526489, -1.346505, -2.593995, -0.771889, 1.570796, 2.097286],accel_mss,speed_ms,0,blend_radius_m)
  movel([0.523400, -1.349714, -2.591876, -0.770799, 1.570796, 2.094196],accel_mss,speed_ms,0,blend_radius_m)
  movel([0.520226, -1.351927, -2.590407, -0.770055, 1.570796, 2.091022],accel_mss,speed_ms,0,blend_radius_m)
  movel([0.517025, -1.353271, -2.589511, -0.769607, 1.570796, 2.087821],accel_mss,speed_ms,0,blend_radius_m)
  speed_ms = 0.003
  movel([0.517025, -1.346591, -2.586414, -0.779384, 1.570796, 2.087821],accel_mss,speed_ms,0,blend_radius_m)
  speed_ms = 0.05
  movel([0.517025, -1.320922, -2.573739, -0.817728, 1.570796, 2.087821],accel_mss,speed_ms,0,blend_radius_m)
  #M_RunCode9
  movel([0.612042, -1.222485, -2.630373, -0.859530, 1.570796, 2.182838],accel_mss,speed_ms,0,blend_radius_m)
  #M_RunCode3
  movel([0.612042, -1.249578, -2.644343, -0.818468, 1.570796, 2.182838],accel_mss,speed_ms,0,blend_radius_m)
  speed_ms = 0.003
  movel([0.612042, -1.256679, -2.647767, -0.807942, 1.570796, 2.182838],accel_mss,speed_ms,0,blend_radius_m)
  speed_ms = 0.007
  movel([0.610850, -1.255352, -2.648485, -0.808552, 1.570796, 2.181646],accel_mss,speed_ms,0,blend_radius_m)
  movel([0.610180, -1.253548, -2.649458, -0.809383, 1.570796, 2.180977],accel_mss,speed_ms,0,blend_radius_m)
  movel([0.609813, -1.251505, -2.650554, -0.810330, 1.570796, 2.180609],accel_mss,speed_ms,0,blend_radius_m)
  movel([0.610746, -1.251259, -2.650686, -0.810444, 1.570796, 2.181542],accel_mss,speed_ms,0,blend_radius_m)
  movel([0.611268, -1.251665, -2.650468, -0.810256, 1.570796, 2.182064],accel_mss,speed_ms,0,blend_radius_m)
  movel([0.611926, -1.252076, -2.650248, -0.810065, 1.570796, 2.182722],accel_mss,speed_ms,0,blend_radius_m)
  movel([0.613261, -1.251850, -2.650369, -0.810170, 1.570796, 2.184057],accel_mss,speed_ms,0,blend_radius_m)
  movel([0.614772, -1.251013, -2.650818, -0.810559, 1.570796, 2.185568],accel_mss,speed_ms,0,blend_radius_m)
  movel([0.616233, -1.249908, -2.651408, -0.811073, 1.570796, 2.187029],accel_mss,speed_ms,0,blend_radius_m)
  movel([0.618237, -1.248311, -2.652258, -0.811820, 1.570796, 2.189033],accel_mss,speed_ms,0,blend_radius_m)
  movel([0.617947, -1.245637, -2.653675, -0.813076, 1.570796, 2.188743],accel_mss,speed_ms,0,blend_radius_m)
  movel([0.616923, -1.243875, -2.654605, -0.813909, 1.570796, 2.187719],accel_mss,speed_ms,0,blend_radius_m)
  movel([0.616065, -1.243468, -2.654819, -0.814102, 1.570796, 2.186862],accel_mss,speed_ms,0,blend_radius_m)
  movel([0.614938, -1.243449, -2.654829, -0.814111, 1.570796, 2.185734],accel_mss,speed_ms,0,blend_radius_m)
  movel([0.613515, -1.243869, -2.654608, -0.813912, 1.570796, 2.184311],accel_mss,speed_ms,0,blend_radius_m)
  movel([0.611773, -1.244776, -2.654130, -0.813483, 1.570796, 2.182570],accel_mss,speed_ms,0,blend_radius_m)
  movel([0.612499, -1.242950, -2.655091, -0.814348, 1.570796, 2.183296],accel_mss,speed_ms,0,blend_radius_m)
  movel([0.613329, -1.241381, -2.655914, -0.815094, 1.570796, 2.184125],accel_mss,speed_ms,0,blend_radius_m)
  movel([0.613825, -1.240829, -2.656203, -0.815357, 1.570796, 2.184622],accel_mss,speed_ms,0,blend_radius_m)
  movel([0.614394, -1.240506, -2.656371, -0.815511, 1.570796, 2.185191],accel_mss,speed_ms,0,blend_radius_m)
  movel([0.615825, -1.240771, -2.656233, -0.815385, 1.570796, 2.186622],accel_mss,speed_ms,0,blend_radius_m)
  movel([0.617921, -1.242529, -2.655312, -0.814548, 1.570796, 2.188718],accel_mss,speed_ms,0,blend_radius_m)
  movel([0.619316, -1.245004, -2.654010, -0.813375, 1.570796, 2.190112],accel_mss,speed_ms,0,blend_radius_m)
  movel([0.619584, -1.246454, -2.653244, -0.812692, 1.570796, 2.190380],accel_mss,speed_ms,0,blend_radius_m)
  movel([0.619474, -1.248016, -2.652415, -0.811958, 1.570796, 2.190270],accel_mss,speed_ms,0,blend_radius_m)
  movel([0.618929, -1.249665, -2.651537, -0.811187, 1.570796, 2.189725],accel_mss,speed_ms,0,blend_radius_m)
  movel([0.617880, -1.251383, -2.650619, -0.810386, 1.570796, 2.188676],accel_mss,speed_ms,0,blend_radius_m)
  movel([0.616504, -1.250348, -2.651173, -0.810868, 1.570796, 2.187301],accel_mss,speed_ms,0,blend_radius_m)
  movel([0.613987, -1.257295, -2.647433, -0.807660, 1.570796, 2.184783],accel_mss,speed_ms,0,blend_radius_m)
  movel([0.612042, -1.256679, -2.647767, -0.807942, 1.570796, 2.182838],accel_mss,speed_ms,0,blend_radius_m)
  speed_ms = 0.003
  movel([0.612042, -1.249578, -2.644343, -0.818468, 1.570796, 2.182838],accel_mss,speed_ms,0,blend_radius_m)
  speed_ms = 0.05
  movel([0.612042, -1.222485, -2.630373, -0.859530, 1.570796, 2.182838],accel_mss,speed_ms,0,blend_radius_m)
  #M_RunCode9
  movel([0.591456, -1.174119, -2.654087, -0.884183, 1.570796, 2.162252],accel_mss,speed_ms,0,blend_radius_m)
  #M_RunCode3
  movel([0.591456, -1.201686, -2.668697, -0.842006, 1.570796, 2.162252],accel_mss,speed_ms,0,blend_radius_m)
  speed_ms = 0.003
  movel([0.591456, -1.208939, -2.672285, -0.831165, 1.570796, 2.162252],accel_mss,speed_ms,0,blend_radius_m)
  speed_ms = 0.007
  movel([0.588359, -1.211205, -2.671180, -0.830004, 1.570796, 2.159155],accel_mss,speed_ms,0,blend_radius_m)
  movel([0.585138, -1.213198, -2.670204, -0.828987, 1.570796, 2.155934],accel_mss,speed_ms,0,blend_radius_m)
  movel([0.581822, -1.214884, -2.669375, -0.828130, 1.570796, 2.152618],accel_mss,speed_ms,0,blend_radius_m)
  movel([0.578445, -1.216225, -2.668713, -0.827451, 1.570796, 2.149242],accel_mss,speed_ms,0,blend_radius_m)
  movel([0.575048, -1.217185, -2.668237, -0.826966, 1.570796, 2.145844],accel_mss,speed_ms,0,blend_radius_m)
  movel([0.573345, -1.217319, -2.668171, -0.826899, 1.570796, 2.144141],accel_mss,speed_ms,0,blend_radius_m)
  movel([0.571660, -1.217172, -2.668244, -0.826973, 1.570796, 2.142456],accel_mss,speed_ms,0,blend_radius_m)
  movel([0.570140, -1.217053, -2.668303, -0.827033, 1.570796, 2.140936],accel_mss,speed_ms,0,blend_radius_m)
  movel([0.568941, -1.217262, -2.668200, -0.826928, 1.570796, 2.139737],accel_mss,speed_ms,0,blend_radius_m)
  movel([0.566873, -1.218693, -2.667489, -0.826207, 1.570796, 2.137669],accel_mss,speed_ms,0,blend_radius_m)
  movel([0.564147, -1.221009, -2.666335, -0.825045, 1.570796, 2.134944],accel_mss,speed_ms,0,blend_radius_m)
  movel([0.561318, -1.223454, -2.665109, -0.823826, 1.570796, 2.132115],accel_mss,speed_ms,0,blend_radius_m)
  movel([0.558932, -1.225284, -2.664188, -0.822917, 1.570796, 2.129728],accel_mss,speed_ms,0,blend_radius_m)
  movel([0.554225, -1.227961, -2.662833, -0.821596, 1.570796, 2.125021],accel_mss,speed_ms,0,blend_radius_m)
  movel([0.550026, -1.229677, -2.661959, -0.820752, 1.570796, 2.120823],accel_mss,speed_ms,0,blend_radius_m)
  movel([0.546288, -1.230531, -2.661524, -0.820334, 1.570796, 2.117084],accel_mss,speed_ms,0,blend_radius_m)
  movel([0.542964, -1.230613, -2.661482, -0.820294, 1.570796, 2.113760],accel_mss,speed_ms,0,blend_radius_m)
  movel([0.540020, -1.230006, -2.661792, -0.820591, 1.570796, 2.110816],accel_mss,speed_ms,0,blend_radius_m)
  movel([0.537407, -1.228804, -2.662404, -0.821181, 1.570796, 2.108203],accel_mss,speed_ms,0,blend_radius_m)
  movel([0.535098, -1.227083, -2.663278, -0.822028, 1.570796, 2.105894],accel_mss,speed_ms,0,blend_radius_m)
  movel([0.533056, -1.224929, -2.664367, -0.823093, 1.570796, 2.103852],accel_mss,speed_ms,0,blend_radius_m)
  movel([0.529627, -1.219666, -2.667005, -0.825718, 1.570796, 2.100423],accel_mss,speed_ms,0,blend_radius_m)
  movel([0.526861, -1.213687, -2.669964, -0.828738, 1.570796, 2.097657],accel_mss,speed_ms,0,blend_radius_m)
  movel([0.522289, -1.202428, -2.675427, -0.834534, 1.570796, 2.093085],accel_mss,speed_ms,0,blend_radius_m)
  movel([0.519671, -1.197902, -2.677583, -0.836904, 1.570796, 2.090467],accel_mss,speed_ms,0,blend_radius_m)
  movel([0.516029, -1.193158, -2.679819, -0.839412, 1.570796, 2.086825],accel_mss,speed_ms,0,blend_radius_m)
  movel([0.511507, -1.188478, -2.682001, -0.841910, 1.570796, 2.082304],accel_mss,speed_ms,0,blend_radius_m)
  movel([0.506261, -1.184167, -2.683990, -0.844232, 1.570796, 2.077057],accel_mss,speed_ms,0,blend_radius_m)
  movel([0.500453, -1.180515, -2.685660, -0.846214, 1.570796, 2.071249],accel_mss,speed_ms,0,blend_radius_m)
  movel([0.494265, -1.177818, -2.686884, -0.847687, 1.570796, 2.065061],accel_mss,speed_ms,0,blend_radius_m)
  movel([0.487893, -1.176356, -2.687544, -0.848489, 1.570796, 2.058690],accel_mss,speed_ms,0,blend_radius_m)
  movel([0.484702, -1.176171, -2.687627, -0.848591, 1.570796, 2.055498],accel_mss,speed_ms,0,blend_radius_m)
  movel([0.481544, -1.176394, -2.687527, -0.848468, 1.570796, 2.052340],accel_mss,speed_ms,0,blend_radius_m)
  movel([0.478145, -1.177057, -2.687228, -0.848105, 1.570796, 2.048941],accel_mss,speed_ms,0,blend_radius_m)
  movel([0.474068, -1.178233, -2.686696, -0.847460, 1.570796, 2.044865],accel_mss,speed_ms,0,blend_radius_m)
  movel([0.469550, -1.179944, -2.685919, -0.846525, 1.570796, 2.040347],accel_mss,speed_ms,0,blend_radius_m)
  movel([0.464822, -1.182215, -2.684884, -0.845290, 1.570796, 2.035619],accel_mss,speed_ms,0,blend_radius_m)
  movel([0.460129, -1.185051, -2.683584, -0.843754, 1.570796, 2.030925],accel_mss,speed_ms,0,blend_radius_m)
  movel([0.455702, -1.188467, -2.682006, -0.841916, 1.570796, 2.026499],accel_mss,speed_ms,0,blend_radius_m)
  movel([0.451783, -1.192465, -2.680144, -0.839780, 1.570796, 2.022579],accel_mss,speed_ms,0,blend_radius_m)
  movel([0.450084, -1.194681, -2.679104, -0.838604, 1.570796, 2.020880],accel_mss,speed_ms,0,blend_radius_m)
  movel([0.448601, -1.197043, -2.677990, -0.837356, 1.570796, 2.019397],accel_mss,speed_ms,0,blend_radius_m)
  movel([0.446977, -1.200728, -2.676239, -0.835422, 1.570796, 2.017773],accel_mss,speed_ms,0,blend_radius_m)
  movel([0.446500, -1.203839, -2.674750, -0.833800, 1.570796, 2.017297],accel_mss,speed_ms,0,blend_radius_m)
  movel([0.447042, -1.206433, -2.673499, -0.832456, 1.570796, 2.017839],accel_mss,speed_ms,0,blend_radius_m)
  movel([0.448472, -1.208568, -2.672465, -0.831356, 1.570796, 2.019268],accel_mss,speed_ms,0,blend_radius_m)
  movel([0.450667, -1.210296, -2.671624, -0.830469, 1.570796, 2.021464],accel_mss,speed_ms,0,blend_radius_m)
  movel([0.453497, -1.211675, -2.670951, -0.829764, 1.570796, 2.024293],accel_mss,speed_ms,0,blend_radius_m)
  movel([0.456848, -1.212751, -2.670423, -0.829214, 1.570796, 2.027644],accel_mss,speed_ms,0,blend_radius_m)
  movel([0.460596, -1.213579, -2.670017, -0.828793, 1.570796, 2.031393],accel_mss,speed_ms,0,blend_radius_m)
  movel([0.468813, -1.214665, -2.669483, -0.828241, 1.570796, 2.039609],accel_mss,speed_ms,0,blend_radius_m)
  movel([0.477206, -1.215290, -2.669175, -0.827925, 1.570796, 2.048002],accel_mss,speed_ms,0,blend_radius_m)
  movel([0.484842, -1.215773, -2.668936, -0.827680, 1.570796, 2.055638],accel_mss,speed_ms,0,blend_radius_m)
  movel([0.490791, -1.216408, -2.668622, -0.827359, 1.570796, 2.061588],accel_mss,speed_ms,0,blend_radius_m)
  movel([0.504732, -1.218734, -2.667469, -0.826186, 1.570796, 2.075528],accel_mss,speed_ms,0,blend_radius_m)
  movel([0.511998, -1.220275, -2.666702, -0.825413, 1.570796, 2.082795],accel_mss,speed_ms,0,blend_radius_m)
  movel([0.517379, -1.221935, -2.665872, -0.824583, 1.570796, 2.088175],accel_mss,speed_ms,0,blend_radius_m)
  movel([0.519222, -1.222939, -2.665368, -0.824082, 1.570796, 2.090019],accel_mss,speed_ms,0,blend_radius_m)
  movel([0.520754, -1.224227, -2.664721, -0.823441, 1.570796, 2.091550],accel_mss,speed_ms,0,blend_radius_m)
  movel([0.522942, -1.227539, -2.663047, -0.821803, 1.570796, 2.093738],accel_mss,speed_ms,0,blend_radius_m)
  movel([0.524046, -1.231652, -2.660951, -0.819786, 1.570796, 2.094843],accel_mss,speed_ms,0,blend_radius_m)
  movel([0.524182, -1.236344, -2.658535, -0.817510, 1.570796, 2.094978],accel_mss,speed_ms,0,blend_radius_m)
  movel([0.523457, -1.241407, -2.655900, -0.815082, 1.570796, 2.094253],accel_mss,speed_ms,0,blend_radius_m)
  movel([0.521980, -1.246636, -2.653147, -0.812606, 1.570796, 2.092776],accel_mss,speed_ms,0,blend_radius_m)
  movel([0.519861, -1.251838, -2.650376, -0.810175, 1.570796, 2.090657],accel_mss,speed_ms,0,blend_radius_m)
  movel([0.517202, -1.256821, -2.647691, -0.807878, 1.570796, 2.087998],accel_mss,speed_ms,0,blend_radius_m)
  movel([0.513213, -1.262651, -2.644511, -0.805227, 1.570796, 2.084010],accel_mss,speed_ms,0,blend_radius_m)
  movel([0.511253, -1.264945, -2.643248, -0.804196, 1.570796, 2.082049],accel_mss,speed_ms,0,blend_radius_m)
  movel([0.509294, -1.266889, -2.642174, -0.803327, 1.570796, 2.080090],accel_mss,speed_ms,0,blend_radius_m)
  movel([0.507324, -1.268518, -2.641269, -0.802602, 1.570796, 2.078120],accel_mss,speed_ms,0,blend_radius_m)
  movel([0.505335, -1.269876, -2.640513, -0.802000, 1.570796, 2.076132],accel_mss,speed_ms,0,blend_radius_m)
  movel([0.501248, -1.271936, -2.639361, -0.801092, 1.570796, 2.072044],accel_mss,speed_ms,0,blend_radius_m)
  movel([0.496932, -1.273384, -2.638548, -0.800457, 1.570796, 2.067729],accel_mss,speed_ms,0,blend_radius_m)
  movel([0.492307, -1.274532, -2.637902, -0.799955, 1.570796, 2.063104],accel_mss,speed_ms,0,blend_radius_m)
  movel([0.481800, -1.277147, -2.636424, -0.798818, 1.570796, 2.052596],accel_mss,speed_ms,0,blend_radius_m)
  movel([0.481250, -1.277333, -2.636319, -0.798738, 1.570796, 2.052047],accel_mss,speed_ms,0,blend_radius_m)
  movel([0.481422, -1.277440, -2.636258, -0.798691, 1.570796, 2.052218],accel_mss,speed_ms,0,blend_radius_m)
  movel([0.483539, -1.277465, -2.636243, -0.798680, 1.570796, 2.054335],accel_mss,speed_ms,0,blend_radius_m)
  movel([0.492250, -1.277066, -2.636469, -0.798853, 1.570796, 2.063046],accel_mss,speed_ms,0,blend_radius_m)
  movel([0.506669, -1.276529, -2.636774, -0.799086, 1.570796, 2.077466],accel_mss,speed_ms,0,blend_radius_m)
  movel([0.498099, -1.280502, -2.634515, -0.797372, 1.570796, 2.068896],accel_mss,speed_ms,0,blend_radius_m)
  movel([0.488583, -1.284504, -2.632219, -0.795666, 1.570796, 2.059379],accel_mss,speed_ms,0,blend_radius_m)
  movel([0.478466, -1.288459, -2.629931, -0.793999, 1.570796, 2.049262],accel_mss,speed_ms,0,blend_radius_m)
  movel([0.468080, -1.292281, -2.627701, -0.792407, 1.570796, 2.038876],accel_mss,speed_ms,0,blend_radius_m)
  movel([0.447854, -1.299150, -2.623645, -0.789594, 1.570796, 2.018650],accel_mss,speed_ms,0,blend_radius_m)
  movel([0.438665, -1.301990, -2.621951, -0.788448, 1.570796, 2.009462],accel_mss,speed_ms,0,blend_radius_m)
  movel([0.430531, -1.304277, -2.620579, -0.787534, 1.570796, 2.001328],accel_mss,speed_ms,0,blend_radius_m)
  movel([0.419111, -1.311715, -2.616068, -0.784605, 1.570796, 1.989907],accel_mss,speed_ms,0,blend_radius_m)
  movel([0.407593, -1.319811, -2.611076, -0.781501, 1.570796, 1.978390],accel_mss,speed_ms,0,blend_radius_m)
  movel([0.384655, -1.336805, -2.600314, -0.775270, 1.570796, 1.955451],accel_mss,speed_ms,0,blend_radius_m)
  movel([0.373383, -1.345165, -2.594876, -0.772348, 1.570796, 1.944179],accel_mss,speed_ms,0,blend_radius_m)
  movel([0.362315, -1.353099, -2.589626, -0.769664, 1.570796, 1.933112],accel_mss,speed_ms,0,blend_radius_m)
  movel([0.351493, -1.360378, -2.584732, -0.767279, 1.570796, 1.922289],accel_mss,speed_ms,0,blend_radius_m)
  movel([0.340941, -1.366779, -2.580368, -0.765243, 1.570796, 1.911737],accel_mss,speed_ms,0,blend_radius_m)
  movel([0.336847, -1.368940, -2.578881, -0.764568, 1.570796, 1.907643],accel_mss,speed_ms,0,blend_radius_m)
  movel([0.332962, -1.370685, -2.577675, -0.764028, 1.570796, 1.903758],accel_mss,speed_ms,0,blend_radius_m)
  movel([0.329303, -1.372019, -2.576752, -0.763619, 1.570796, 1.900099],accel_mss,speed_ms,0,blend_radius_m)
  movel([0.325892, -1.372944, -2.576109, -0.763336, 1.570796, 1.896688],accel_mss,speed_ms,0,blend_radius_m)
  movel([0.322744, -1.373466, -2.575746, -0.763177, 1.570796, 1.893540],accel_mss,speed_ms,0,blend_radius_m)
  movel([0.319880, -1.373584, -2.575664, -0.763141, 1.570796, 1.890677],accel_mss,speed_ms,0,blend_radius_m)
  movel([0.317326, -1.373299, -2.575862, -0.763228, 1.570796, 1.888122],accel_mss,speed_ms,0,blend_radius_m)
  movel([0.315102, -1.372611, -2.576340, -0.763438, 1.570796, 1.885898],accel_mss,speed_ms,0,blend_radius_m)
  movel([0.313228, -1.371518, -2.577098, -0.763772, 1.570796, 1.884024],accel_mss,speed_ms,0,blend_radius_m)
  movel([0.311733, -1.370020, -2.578136, -0.764234, 1.570796, 1.882529],accel_mss,speed_ms,0,blend_radius_m)
  movel([0.310641, -1.368110, -2.579452, -0.764826, 1.570796, 1.881438],accel_mss,speed_ms,0,blend_radius_m)
  movel([0.309977, -1.365788, -2.581047, -0.765554, 1.570796, 1.880773],accel_mss,speed_ms,0,blend_radius_m)
  movel([0.309771, -1.363045, -2.582921, -0.766423, 1.570796, 1.880567],accel_mss,speed_ms,0,blend_radius_m)
  movel([0.310052, -1.359877, -2.585071, -0.767441, 1.570796, 1.880849],accel_mss,speed_ms,0,blend_radius_m)
  movel([0.310849, -1.356277, -2.587499, -0.768614, 1.570796, 1.881645],accel_mss,speed_ms,0,blend_radius_m)
  movel([0.312198, -1.352239, -2.590199, -0.769951, 1.570796, 1.882995],accel_mss,speed_ms,0,blend_radius_m)
  movel([0.315388, -1.353373, -2.589443, -0.769573, 1.570796, 1.886184],accel_mss,speed_ms,0,blend_radius_m)
  movel([0.317012, -1.353821, -2.589144, -0.769424, 1.570796, 1.887808],accel_mss,speed_ms,0,blend_radius_m)
  movel([0.318807, -1.353826, -2.589140, -0.769423, 1.570796, 1.889604],accel_mss,speed_ms,0,blend_radius_m)
  movel([0.320368, -1.353349, -2.589459, -0.769581, 1.570796, 1.891164],accel_mss,speed_ms,0,blend_radius_m)
  movel([0.322310, -1.352386, -2.590101, -0.769902, 1.570796, 1.893106],accel_mss,speed_ms,0,blend_radius_m)
  movel([0.327139, -1.349239, -2.592191, -0.770959, 1.570796, 1.897935],accel_mss,speed_ms,0,blend_radius_m)
  movel([0.332894, -1.344852, -2.595081, -0.772456, 1.570796, 1.903690],accel_mss,speed_ms,0,blend_radius_m)
  movel([0.339162, -1.339703, -2.598440, -0.774246, 1.570796, 1.909959],accel_mss,speed_ms,0,blend_radius_m)
  movel([0.351512, -1.329039, -2.605281, -0.778069, 1.570796, 1.922308],accel_mss,speed_ms,0,blend_radius_m)
  movel([0.360542, -1.321245, -2.610184, -0.780961, 1.570796, 1.931338],accel_mss,speed_ms,0,blend_radius_m)
  movel([0.368674, -1.314968, -2.614073, -0.783348, 1.570796, 1.939470],accel_mss,speed_ms,0,blend_radius_m)
  movel([0.376896, -1.308658, -2.617931, -0.785800, 1.570796, 1.947692],accel_mss,speed_ms,0,blend_radius_m)
  movel([0.360318, -1.312132, -2.615813, -0.784444, 1.570796, 1.931114],accel_mss,speed_ms,0,blend_radius_m)
  movel([0.351766, -1.313610, -2.614908, -0.783871, 1.570796, 1.922562],accel_mss,speed_ms,0,blend_radius_m)
  movel([0.343643, -1.314328, -2.614467, -0.783594, 1.570796, 1.914440],accel_mss,speed_ms,0,blend_radius_m)
  movel([0.339880, -1.314262, -2.614507, -0.783620, 1.570796, 1.910677],accel_mss,speed_ms,0,blend_radius_m)
  movel([0.336389, -1.313837, -2.614769, -0.783784, 1.570796, 1.907185],accel_mss,speed_ms,0,blend_radius_m)
  movel([0.333222, -1.312993, -2.615286, -0.784110, 1.570796, 1.904018],accel_mss,speed_ms,0,blend_radius_m)
  movel([0.330436, -1.311668, -2.616097, -0.784624, 1.570796, 1.901232],accel_mss,speed_ms,0,blend_radius_m)
  movel([0.328086, -1.309807, -2.617232, -0.785350, 1.570796, 1.898882],accel_mss,speed_ms,0,blend_radius_m)
  movel([0.326231, -1.307337, -2.618732, -0.786320, 1.570796, 1.897027],accel_mss,speed_ms,0,blend_radius_m)
  movel([0.324928, -1.304198, -2.620626, -0.787565, 1.570796, 1.895724],accel_mss,speed_ms,0,blend_radius_m)
  movel([0.324237, -1.300315, -2.622951, -0.789123, 1.570796, 1.895034],accel_mss,speed_ms,0,blend_radius_m)
  movel([0.324402, -1.295276, -2.625940, -0.791173, 1.570796, 1.895199],accel_mss,speed_ms,0,blend_radius_m)
  movel([0.325635, -1.289753, -2.629178, -0.793458, 1.570796, 1.896431],accel_mss,speed_ms,0,blend_radius_m)
  movel([0.327860, -1.283913, -2.632560, -0.795916, 1.570796, 1.898656],accel_mss,speed_ms,0,blend_radius_m)
  movel([0.330982, -1.277944, -2.635971, -0.798473, 1.570796, 1.901779],accel_mss,speed_ms,0,blend_radius_m)
  movel([0.334915, -1.272036, -2.639305, -0.801048, 1.570796, 1.905711],accel_mss,speed_ms,0,blend_radius_m)
  movel([0.339561, -1.266390, -2.642450, -0.803549, 1.570796, 1.910357],accel_mss,speed_ms,0,blend_radius_m)
  movel([0.344810, -1.261214, -2.645299, -0.805877, 1.570796, 1.915606],accel_mss,speed_ms,0,blend_radius_m)
  movel([0.350551, -1.256727, -2.647742, -0.807921, 1.570796, 1.921348],accel_mss,speed_ms,0,blend_radius_m)
  movel([0.353841, -1.254968, -2.648692, -0.808728, 1.570796, 1.924637],accel_mss,speed_ms,0,blend_radius_m)
  movel([0.357509, -1.253715, -2.649367, -0.809306, 1.570796, 1.928305],accel_mss,speed_ms,0,blend_radius_m)
  movel([0.360374, -1.253441, -2.649515, -0.809433, 1.570796, 1.931170],accel_mss,speed_ms,0,blend_radius_m)
  movel([0.361138, -1.253812, -2.649315, -0.809261, 1.570796, 1.931934],accel_mss,speed_ms,0,blend_radius_m)
  movel([0.361259, -1.254595, -2.648894, -0.808900, 1.570796, 1.932055],accel_mss,speed_ms,0,blend_radius_m)
  movel([0.358364, -1.255534, -2.648387, -0.808468, 1.570796, 1.929161],accel_mss,speed_ms,0,blend_radius_m)
  movel([0.355887, -1.256629, -2.647794, -0.807965, 1.570796, 1.926683],accel_mss,speed_ms,0,blend_radius_m)
  movel([0.353810, -1.257855, -2.647130, -0.807404, 1.570796, 1.924607],accel_mss,speed_ms,0,blend_radius_m)
  movel([0.352126, -1.259180, -2.646409, -0.806800, 1.570796, 1.922923],accel_mss,speed_ms,0,blend_radius_m)
  movel([0.350820, -1.260578, -2.645646, -0.806165, 1.570796, 1.921617],accel_mss,speed_ms,0,blend_radius_m)
  movel([0.349874, -1.262022, -2.644856, -0.805511, 1.570796, 1.920671],accel_mss,speed_ms,0,blend_radius_m)
  movel([0.349276, -1.263485, -2.644053, -0.804852, 1.570796, 1.920073],accel_mss,speed_ms,0,blend_radius_m)
  movel([0.349011, -1.264947, -2.643247, -0.804195, 1.570796, 1.919808],accel_mss,speed_ms,0,blend_radius_m)
  movel([0.349414, -1.267755, -2.641693, -0.802941, 1.570796, 1.920210],accel_mss,speed_ms,0,blend_radius_m)
  movel([0.350963, -1.270260, -2.640299, -0.801831, 1.570796, 1.921759],accel_mss,speed_ms,0,blend_radius_m)
  movel([0.353545, -1.272265, -2.639176, -0.800947, 1.570796, 1.924341],accel_mss,speed_ms,0,blend_radius_m)
  movel([0.357041, -1.273591, -2.638432, -0.800366, 1.570796, 1.927837],accel_mss,speed_ms,0,blend_radius_m)
  movel([0.359470, -1.273903, -2.638256, -0.800230, 1.570796, 1.930267],accel_mss,speed_ms,0,blend_radius_m)
  movel([0.362592, -1.273890, -2.638264, -0.800236, 1.570796, 1.933388],accel_mss,speed_ms,0,blend_radius_m)
  movel([0.370536, -1.273052, -2.638735, -0.800602, 1.570796, 1.941333],accel_mss,speed_ms,0,blend_radius_m)
  movel([0.380143, -1.271395, -2.639664, -0.801330, 1.570796, 1.950940],accel_mss,speed_ms,0,blend_radius_m)
  movel([0.390687, -1.269207, -2.640886, -0.802297, 1.570796, 1.961483],accel_mss,speed_ms,0,blend_radius_m)
  movel([0.411673, -1.264310, -2.643599, -0.804481, 1.570796, 1.982469],accel_mss,speed_ms,0,blend_radius_m)
  movel([0.427610, -1.260313, -2.645791, -0.806285, 1.570796, 1.998406],accel_mss,speed_ms,0,blend_radius_m)
  movel([0.435645, -1.258294, -2.646891, -0.807204, 1.570796, 2.006442],accel_mss,speed_ms,0,blend_radius_m)
  movel([0.440000, -1.257068, -2.647557, -0.807765, 1.570796, 2.010796],accel_mss,speed_ms,0,blend_radius_m)
  movel([0.443348, -1.255835, -2.648224, -0.808330, 1.570796, 2.014144],accel_mss,speed_ms,0,blend_radius_m)
  movel([0.444277, -1.255304, -2.648511, -0.808574, 1.570796, 2.015073],accel_mss,speed_ms,0,blend_radius_m)
  movel([0.444664, -1.254829, -2.648767, -0.808792, 1.570796, 2.015460],accel_mss,speed_ms,0,blend_radius_m)
  movel([0.444259, -1.253781, -2.649332, -0.809276, 1.570796, 2.015055],accel_mss,speed_ms,0,blend_radius_m)
  movel([0.441834, -1.251674, -2.650463, -0.810251, 1.570796, 2.012630],accel_mss,speed_ms,0,blend_radius_m)
  movel([0.438704, -1.250151, -2.651278, -0.810960, 1.570796, 2.009501],accel_mss,speed_ms,0,blend_radius_m)
  movel([0.431646, -1.247295, -2.652798, -0.812296, 1.570796, 2.002442],accel_mss,speed_ms,0,blend_radius_m)
  movel([0.428373, -1.245163, -2.653926, -0.813300, 1.570796, 1.999170],accel_mss,speed_ms,0,blend_radius_m)
  movel([0.425709, -1.242013, -2.655583, -0.814793, 1.570796, 1.996505],accel_mss,speed_ms,0,blend_radius_m)
  movel([0.424705, -1.239924, -2.656676, -0.815790, 1.570796, 1.995501],accel_mss,speed_ms,0,blend_radius_m)
  movel([0.423981, -1.237416, -2.657980, -0.816993, 1.570796, 1.994777],accel_mss,speed_ms,0,blend_radius_m)
  movel([0.423574, -1.234437, -2.659520, -0.818432, 1.570796, 1.994370],accel_mss,speed_ms,0,blend_radius_m)
  movel([0.423533, -1.230923, -2.661324, -0.820142, 1.570796, 1.994329],accel_mss,speed_ms,0,blend_radius_m)
  movel([0.424200, -1.225986, -2.663833, -0.822570, 1.570796, 1.994997],accel_mss,speed_ms,0,blend_radius_m)
  movel([0.425746, -1.221017, -2.666331, -0.825041, 1.570796, 1.996543],accel_mss,speed_ms,0,blend_radius_m)
  movel([0.428072, -1.216036, -2.668806, -0.827547, 1.570796, 1.998868],accel_mss,speed_ms,0,blend_radius_m)
  movel([0.431076, -1.211066, -2.671248, -0.830075, 1.570796, 2.001872],accel_mss,speed_ms,0,blend_radius_m)
  movel([0.434656, -1.206129, -2.673646, -0.832614, 1.570796, 2.005452],accel_mss,speed_ms,0,blend_radius_m)
  movel([0.438707, -1.201247, -2.675991, -0.835151, 1.570796, 2.009504],accel_mss,speed_ms,0,blend_radius_m)
  movel([0.443125, -1.196449, -2.678270, -0.837669, 1.570796, 2.013921],accel_mss,speed_ms,0,blend_radius_m)
  movel([0.447799, -1.191757, -2.680475, -0.840157, 1.570796, 2.018595],accel_mss,speed_ms,0,blend_radius_m)
  movel([0.457028, -1.183464, -2.684313, -0.844613, 1.570796, 2.027824],accel_mss,speed_ms,0,blend_radius_m)
  movel([0.465504, -1.176943, -2.687279, -0.848167, 1.570796, 2.036300],accel_mss,speed_ms,0,blend_radius_m)
  movel([0.472808, -1.172123, -2.689443, -0.850823, 1.570796, 2.043604],accel_mss,speed_ms,0,blend_radius_m)
  movel([0.478525, -1.168909, -2.690872, -0.852608, 1.570796, 2.049321],accel_mss,speed_ms,0,blend_radius_m)
  movel([0.486982, -1.165142, -2.692534, -0.854714, 1.570796, 2.057778],accel_mss,speed_ms,0,blend_radius_m)
  movel([0.495103, -1.162621, -2.693637, -0.856131, 1.570796, 2.065899],accel_mss,speed_ms,0,blend_radius_m)
  movel([0.502783, -1.161328, -2.694201, -0.856860, 1.570796, 2.073580],accel_mss,speed_ms,0,blend_radius_m)
  movel([0.509918, -1.161234, -2.694241, -0.856913, 1.570796, 2.080715],accel_mss,speed_ms,0,blend_radius_m)
  movel([0.516406, -1.162302, -2.693776, -0.856310, 1.570796, 2.087202],accel_mss,speed_ms,0,blend_radius_m)
  movel([0.522160, -1.164477, -2.692825, -0.855087, 1.570796, 2.092957],accel_mss,speed_ms,0,blend_radius_m)
  movel([0.527100, -1.167701, -2.691406, -0.853281, 1.570796, 2.097896],accel_mss,speed_ms,0,blend_radius_m)
  movel([0.531147, -1.171908, -2.689539, -0.850943, 1.570796, 2.101944],accel_mss,speed_ms,0,blend_radius_m)
  movel([0.533972, -1.176476, -2.687490, -0.848423, 1.570796, 2.104769],accel_mss,speed_ms,0,blend_radius_m)
  movel([0.536246, -1.181445, -2.685236, -0.845708, 1.570796, 2.107042],accel_mss,speed_ms,0,blend_radius_m)
  movel([0.538383, -1.186394, -2.682965, -0.843030, 1.570796, 2.109179],accel_mss,speed_ms,0,blend_radius_m)
  movel([0.540780, -1.190926, -2.680863, -0.840600, 1.570796, 2.111576],accel_mss,speed_ms,0,blend_radius_m)
  movel([0.543836, -1.194654, -2.679117, -0.838618, 1.570796, 2.114632],accel_mss,speed_ms,0,blend_radius_m)
  movel([0.545735, -1.196100, -2.678435, -0.837854, 1.570796, 2.116532],accel_mss,speed_ms,0,blend_radius_m)
  movel([0.547946, -1.197211, -2.677910, -0.837268, 1.570796, 2.118742],accel_mss,speed_ms,0,blend_radius_m)
  movel([0.550519, -1.197931, -2.677569, -0.836889, 1.570796, 2.121316],accel_mss,speed_ms,0,blend_radius_m)
  movel([0.553510, -1.198224, -2.677430, -0.836735, 1.570796, 2.124306],accel_mss,speed_ms,0,blend_radius_m)
  movel([0.556965, -1.198040, -2.677518, -0.836832, 1.570796, 2.127761],accel_mss,speed_ms,0,blend_radius_m)
  movel([0.560936, -1.197335, -2.677852, -0.837203, 1.570796, 2.131732],accel_mss,speed_ms,0,blend_radius_m)
  movel([0.564567, -1.196167, -2.678403, -0.837818, 1.570796, 2.135363],accel_mss,speed_ms,0,blend_radius_m)
  movel([0.567769, -1.194505, -2.679187, -0.838697, 1.570796, 2.138566],accel_mss,speed_ms,0,blend_radius_m)
  movel([0.570539, -1.192442, -2.680155, -0.839793, 1.570796, 2.141336],accel_mss,speed_ms,0,blend_radius_m)
  movel([0.572877, -1.190070, -2.681262, -0.841057, 1.570796, 2.143673],accel_mss,speed_ms,0,blend_radius_m)
  movel([0.574767, -1.187494, -2.682457, -0.842438, 1.570796, 2.145563],accel_mss,speed_ms,0,blend_radius_m)
  movel([0.576199, -1.184810, -2.683695, -0.843884, 1.570796, 2.146996],accel_mss,speed_ms,0,blend_radius_m)
  movel([0.577167, -1.182123, -2.684926, -0.845339, 1.570796, 2.147963],accel_mss,speed_ms,0,blend_radius_m)
  movel([0.577656, -1.179539, -2.686104, -0.846746, 1.570796, 2.148452],accel_mss,speed_ms,0,blend_radius_m)
  movel([0.577647, -1.177168, -2.687177, -0.848043, 1.570796, 2.148443],accel_mss,speed_ms,0,blend_radius_m)
  movel([0.577132, -1.175122, -2.688099, -0.849168, 1.570796, 2.147928],accel_mss,speed_ms,0,blend_radius_m)
  movel([0.576096, -1.173511, -2.688822, -0.850056, 1.570796, 2.146893],accel_mss,speed_ms,0,blend_radius_m)
  movel([0.574529, -1.172448, -2.689298, -0.850643, 1.570796, 2.145325],accel_mss,speed_ms,0,blend_radius_m)
  movel([0.572421, -1.172043, -2.689478, -0.850867, 1.570796, 2.143217],accel_mss,speed_ms,0,blend_radius_m)
  movel([0.569766, -1.172407, -2.689316, -0.850666, 1.570796, 2.140563],accel_mss,speed_ms,0,blend_radius_m)
  movel([0.566559, -1.173646, -2.688761, -0.849981, 1.570796, 2.137355],accel_mss,speed_ms,0,blend_radius_m)
  movel([0.562802, -1.175864, -2.687765, -0.848759, 1.570796, 2.133598],accel_mss,speed_ms,0,blend_radius_m)
  movel([0.564785, -1.176270, -2.687583, -0.848536, 1.570796, 2.135582],accel_mss,speed_ms,0,blend_radius_m)
  movel([0.566165, -1.177085, -2.687215, -0.848089, 1.570796, 2.136961],accel_mss,speed_ms,0,blend_radius_m)
  movel([0.566937, -1.178246, -2.686690, -0.847453, 1.570796, 2.137733],accel_mss,speed_ms,0,blend_radius_m)
  movel([0.567097, -1.179689, -2.686035, -0.846664, 1.570796, 2.137893],accel_mss,speed_ms,0,blend_radius_m)
  movel([0.566633, -1.181357, -2.685276, -0.845756, 1.570796, 2.137429],accel_mss,speed_ms,0,blend_radius_m)
  movel([0.565551, -1.183185, -2.684441, -0.844763, 1.570796, 2.136347],accel_mss,speed_ms,0,blend_radius_m)
  movel([0.563839, -1.185112, -2.683556, -0.843721, 1.570796, 2.134635],accel_mss,speed_ms,0,blend_radius_m)
  movel([0.561493, -1.187090, -2.682644, -0.842655, 1.570796, 2.132289],accel_mss,speed_ms,0,blend_radius_m)
  movel([0.557225, -1.189752, -2.681409, -0.841227, 1.570796, 2.128022],accel_mss,speed_ms,0,blend_radius_m)
  movel([0.553383, -1.191179, -2.680745, -0.840465, 1.570796, 2.124179],accel_mss,speed_ms,0,blend_radius_m)
  movel([0.549982, -1.191502, -2.680594, -0.840293, 1.570796, 2.120778],accel_mss,speed_ms,0,blend_radius_m)
  movel([0.547041, -1.190838, -2.680904, -0.840647, 1.570796, 2.117837],accel_mss,speed_ms,0,blend_radius_m)
  movel([0.544592, -1.189297, -2.681621, -0.841471, 1.570796, 2.115388],accel_mss,speed_ms,0,blend_radius_m)
  movel([0.542665, -1.186993, -2.682689, -0.842708, 1.570796, 2.113461],accel_mss,speed_ms,0,blend_radius_m)
  movel([0.541298, -1.184022, -2.684057, -0.844310, 1.570796, 2.112095],accel_mss,speed_ms,0,blend_radius_m)
  movel([0.540524, -1.180498, -2.685668, -0.846224, 1.570796, 2.111321],accel_mss,speed_ms,0,blend_radius_m)
  movel([0.540393, -1.176522, -2.687469, -0.848398, 1.570796, 2.111189],accel_mss,speed_ms,0,blend_radius_m)
  movel([0.540940, -1.172199, -2.689409, -0.850781, 1.570796, 2.111737],accel_mss,speed_ms,0,blend_radius_m)
  movel([0.542216, -1.167638, -2.691434, -0.853317, 1.570796, 2.113013],accel_mss,speed_ms,0,blend_radius_m)
  movel([0.544265, -1.162953, -2.693492, -0.855944, 1.570796, 2.115062],accel_mss,speed_ms,0,blend_radius_m)
  movel([0.547138, -1.158257, -2.695532, -0.858600, 1.570796, 2.117935],accel_mss,speed_ms,0,blend_radius_m)
  movel([0.550870, -1.153678, -2.697500, -0.861211, 1.570796, 2.121666],accel_mss,speed_ms,0,blend_radius_m)
  movel([0.555507, -1.149347, -2.699342, -0.863700, 1.570796, 2.126303],accel_mss,speed_ms,0,blend_radius_m)
  movel([0.561079, -1.145401, -2.701003, -0.865985, 1.570796, 2.131875],accel_mss,speed_ms,0,blend_radius_m)
  movel([0.565226, -1.143044, -2.701988, -0.867357, 1.570796, 2.136022],accel_mss,speed_ms,0,blend_radius_m)
  movel([0.569346, -1.141066, -2.702811, -0.868512, 1.570796, 2.140142],accel_mss,speed_ms,0,blend_radius_m)
  movel([0.573400, -1.139478, -2.703468, -0.869443, 1.570796, 2.144196],accel_mss,speed_ms,0,blend_radius_m)
  movel([0.577358, -1.138281, -2.703962, -0.870146, 1.570796, 2.148154],accel_mss,speed_ms,0,blend_radius_m)
  movel([0.581178, -1.137489, -2.704288, -0.870612, 1.570796, 2.151974],accel_mss,speed_ms,0,blend_radius_m)
  movel([0.584826, -1.137105, -2.704446, -0.870838, 1.570796, 2.155622],accel_mss,speed_ms,0,blend_radius_m)
  movel([0.588269, -1.137134, -2.704434, -0.870821, 1.570796, 2.159065],accel_mss,speed_ms,0,blend_radius_m)
  movel([0.591474, -1.137578, -2.704252, -0.870560, 1.570796, 2.162271],accel_mss,speed_ms,0,blend_radius_m)
  movel([0.594401, -1.138446, -2.703894, -0.870049, 1.570796, 2.165197],accel_mss,speed_ms,0,blend_radius_m)
  movel([0.597024, -1.139731, -2.703364, -0.869295, 1.570796, 2.167820],accel_mss,speed_ms,0,blend_radius_m)
  movel([0.599307, -1.141435, -2.702658, -0.868296, 1.570796, 2.170103],accel_mss,speed_ms,0,blend_radius_m)
  movel([0.601221, -1.143559, -2.701774, -0.867056, 1.570796, 2.172018],accel_mss,speed_ms,0,blend_radius_m)
  movel([0.602739, -1.146096, -2.700712, -0.865581, 1.570796, 2.173536],accel_mss,speed_ms,0,blend_radius_m)
  movel([0.603829, -1.149044, -2.699470, -0.863875, 1.570796, 2.174626],accel_mss,speed_ms,0,blend_radius_m)
  movel([0.604466, -1.152395, -2.698048, -0.861947, 1.570796, 2.175262],accel_mss,speed_ms,0,blend_radius_m)
  movel([0.604628, -1.156147, -2.696442, -0.859800, 1.570796, 2.175424],accel_mss,speed_ms,0,blend_radius_m)
  movel([0.603835, -1.160294, -2.694650, -0.857445, 1.570796, 2.174631],accel_mss,speed_ms,0,blend_radius_m)
  movel([0.602201, -1.165017, -2.692588, -0.854784, 1.570796, 2.172997],accel_mss,speed_ms,0,blend_radius_m)
  movel([0.600598, -1.169104, -2.690785, -0.852499, 1.570796, 2.171394],accel_mss,speed_ms,0,blend_radius_m)
  movel([0.599873, -1.171394, -2.689768, -0.851227, 1.570796, 2.170670],accel_mss,speed_ms,0,blend_radius_m)
  movel([0.600660, -1.172529, -2.689261, -0.850598, 1.570796, 2.171457],accel_mss,speed_ms,0,blend_radius_m)
  movel([0.602471, -1.173882, -2.688656, -0.849851, 1.570796, 2.173267],accel_mss,speed_ms,0,blend_radius_m)
  movel([0.604468, -1.175370, -2.687988, -0.849031, 1.570796, 2.175264],accel_mss,speed_ms,0,blend_radius_m)
  movel([0.605816, -1.176909, -2.687294, -0.848186, 1.570796, 2.176613],accel_mss,speed_ms,0,blend_radius_m)
  movel([0.606776, -1.179604, -2.686074, -0.846711, 1.570796, 2.177572],accel_mss,speed_ms,0,blend_radius_m)
  movel([0.607148, -1.182477, -2.684765, -0.845148, 1.570796, 2.177944],accel_mss,speed_ms,0,blend_radius_m)
  movel([0.606981, -1.185479, -2.683387, -0.843523, 1.570796, 2.177777],accel_mss,speed_ms,0,blend_radius_m)
  movel([0.606318, -1.188563, -2.681962, -0.841864, 1.570796, 2.177115],accel_mss,speed_ms,0,blend_radius_m)
  movel([0.605205, -1.191687, -2.680507, -0.840194, 1.570796, 2.176001],accel_mss,speed_ms,0,blend_radius_m)
  movel([0.603685, -1.194809, -2.679044, -0.838536, 1.570796, 2.174481],accel_mss,speed_ms,0,blend_radius_m)
  movel([0.601801, -1.197884, -2.677592, -0.836914, 1.570796, 2.172598],accel_mss,speed_ms,0,blend_radius_m)
  movel([0.599596, -1.200872, -2.676170, -0.835347, 1.570796, 2.170392],accel_mss,speed_ms,0,blend_radius_m)
  movel([0.597110, -1.203736, -2.674799, -0.833854, 1.570796, 2.167907],accel_mss,speed_ms,0,blend_radius_m)
  movel([0.594383, -1.206440, -2.673496, -0.832453, 1.570796, 2.165179],accel_mss,speed_ms,0,blend_radius_m)
  movel([0.591456, -1.208939, -2.672285, -0.831165, 1.570796, 2.162252],accel_mss,speed_ms,0,blend_radius_m)
  speed_ms = 0.003
  movel([0.591456, -1.201686, -2.668697, -0.842006, 1.570796, 2.162252],accel_mss,speed_ms,0,blend_radius_m)
  speed_ms = 0.05
  movel([0.591456, -1.174119, -2.654087, -0.884183, 1.570796, 2.162252],accel_mss,speed_ms,0,blend_radius_m)
  #M_RunCode9
  movel([0.610750, -1.173087, -2.654565, -0.884737, 1.570796, 2.181547],accel_mss,speed_ms,0,blend_radius_m)
  #M_RunCode3
  movel([0.610750, -1.200662, -2.669189, -0.842538, 1.570796, 2.181547],accel_mss,speed_ms,0,blend_radius_m)
  speed_ms = 0.003
  movel([0.610750, -1.207918, -2.672780, -0.831690, 1.570796, 2.181547],accel_mss,speed_ms,0,blend_radius_m)
  speed_ms = 0.007
  movel([0.611982, -1.205326, -2.674034, -0.833029, 1.570796, 2.182779],accel_mss,speed_ms,0,blend_radius_m)
  movel([0.615148, -1.200057, -2.676559, -0.835773, 1.570796, 2.185945],accel_mss,speed_ms,0,blend_radius_m)
  movel([0.618029, -1.194878, -2.679011, -0.838500, 1.570796, 2.188825],accel_mss,speed_ms,0,blend_radius_m)
  movel([0.618889, -1.192407, -2.680171, -0.839811, 1.570796, 2.189686],accel_mss,speed_ms,0,blend_radius_m)
  movel([0.619108, -1.190062, -2.681265, -0.841062, 1.570796, 2.189904],accel_mss,speed_ms,0,blend_radius_m)
  movel([0.619540, -1.191482, -2.680603, -0.840304, 1.570796, 2.190336],accel_mss,speed_ms,0,blend_radius_m)
  movel([0.619683, -1.194404, -2.679234, -0.838751, 1.570796, 2.190480],accel_mss,speed_ms,0,blend_radius_m)
  movel([0.619057, -1.197378, -2.677831, -0.837180, 1.570796, 2.189854],accel_mss,speed_ms,0,blend_radius_m)
  movel([0.617905, -1.200392, -2.676399, -0.835598, 1.570796, 2.188701],accel_mss,speed_ms,0,blend_radius_m)
  movel([0.616462, -1.203425, -2.674948, -0.834015, 1.570796, 2.187258],accel_mss,speed_ms,0,blend_radius_m)
  movel([0.613647, -1.209496, -2.672014, -0.830879, 1.570796, 2.184443],accel_mss,speed_ms,0,blend_radius_m)
  movel([0.612739, -1.212503, -2.670545, -0.829341, 1.570796, 2.183535],accel_mss,speed_ms,0,blend_radius_m)
  movel([0.612469, -1.215472, -2.669085, -0.827832, 1.570796, 2.183266],accel_mss,speed_ms,0,blend_radius_m)
  movel([0.612864, -1.218518, -2.667576, -0.826295, 1.570796, 2.183661],accel_mss,speed_ms,0,blend_radius_m)
  movel([0.613252, -1.220047, -2.666815, -0.825527, 1.570796, 2.184048],accel_mss,speed_ms,0,blend_radius_m)
  movel([0.613722, -1.220773, -2.666453, -0.825163, 1.570796, 2.184518],accel_mss,speed_ms,0,blend_radius_m)
  movel([0.615419, -1.220175, -2.666751, -0.825463, 1.570796, 2.186216],accel_mss,speed_ms,0,blend_radius_m)
  movel([0.616806, -1.219753, -2.666962, -0.825674, 1.570796, 2.187602],accel_mss,speed_ms,0,blend_radius_m)
  movel([0.618157, -1.219600, -2.667038, -0.825751, 1.570796, 2.188953],accel_mss,speed_ms,0,blend_radius_m)
  movel([0.620546, -1.219954, -2.666861, -0.825574, 1.570796, 2.191342],accel_mss,speed_ms,0,blend_radius_m)
  movel([0.622088, -1.220655, -2.666512, -0.825222, 1.570796, 2.192885],accel_mss,speed_ms,0,blend_radius_m)
  movel([0.622966, -1.221660, -2.666009, -0.824720, 1.570796, 2.193763],accel_mss,speed_ms,0,blend_radius_m)
  movel([0.623363, -1.222920, -2.665377, -0.824091, 1.570796, 2.194160],accel_mss,speed_ms,0,blend_radius_m)
  movel([0.623428, -1.226047, -2.663803, -0.822540, 1.570796, 2.194225],accel_mss,speed_ms,0,blend_radius_m)
  movel([0.623723, -1.229689, -2.661954, -0.820746, 1.570796, 2.194519],accel_mss,speed_ms,0,blend_radius_m)
  movel([0.625032, -1.234082, -2.659703, -0.818604, 1.570796, 2.195828],accel_mss,speed_ms,0,blend_radius_m)
  movel([0.626531, -1.238312, -2.657515, -0.816562, 1.570796, 2.197328],accel_mss,speed_ms,0,blend_radius_m)
  movel([0.627764, -1.242674, -2.655236, -0.814479, 1.570796, 2.198560],accel_mss,speed_ms,0,blend_radius_m)
  movel([0.628292, -1.247444, -2.652719, -0.812226, 1.570796, 2.199088],accel_mss,speed_ms,0,blend_radius_m)
  movel([0.628109, -1.250233, -2.651234, -0.810922, 1.570796, 2.198906],accel_mss,speed_ms,0,blend_radius_m)
  movel([0.627596, -1.253116, -2.649690, -0.809583, 1.570796, 2.198393],accel_mss,speed_ms,0,blend_radius_m)
  movel([0.625914, -1.259024, -2.646494, -0.806871, 1.570796, 2.196710],accel_mss,speed_ms,0,blend_radius_m)
  movel([0.623924, -1.264893, -2.643277, -0.804219, 1.570796, 2.194720],accel_mss,speed_ms,0,blend_radius_m)
  movel([0.622275, -1.270457, -2.640188, -0.801743, 1.570796, 2.193072],accel_mss,speed_ms,0,blend_radius_m)
  movel([0.620692, -1.279329, -2.635184, -0.797876, 1.570796, 2.191489],accel_mss,speed_ms,0,blend_radius_m)
  movel([0.620124, -1.283073, -2.633043, -0.796274, 1.570796, 2.190921],accel_mss,speed_ms,0,blend_radius_m)
  movel([0.619349, -1.286652, -2.630979, -0.794758, 1.570796, 2.190145],accel_mss,speed_ms,0,blend_radius_m)
  movel([0.618108, -1.290284, -2.628869, -0.793237, 1.570796, 2.188904],accel_mss,speed_ms,0,blend_radius_m)
  movel([0.616143, -1.294177, -2.626587, -0.791625, 1.570796, 2.186940],accel_mss,speed_ms,0,blend_radius_m)
  movel([0.613203, -1.298542, -2.624007, -0.789841, 1.570796, 2.184000],accel_mss,speed_ms,0,blend_radius_m)
  movel([0.609053, -1.303576, -2.621000, -0.787813, 1.570796, 2.179849],accel_mss,speed_ms,0,blend_radius_m)
  movel([0.605359, -1.307458, -2.618659, -0.786273, 1.570796, 2.176156],accel_mss,speed_ms,0,blend_radius_m)
  movel([0.601699, -1.310781, -2.616639, -0.784969, 1.570796, 2.172495],accel_mss,speed_ms,0,blend_radius_m)
  movel([0.598075, -1.313585, -2.614923, -0.783881, 1.570796, 2.168872],accel_mss,speed_ms,0,blend_radius_m)
  movel([0.594488, -1.315900, -2.613499, -0.782990, 1.570796, 2.165284],accel_mss,speed_ms,0,blend_radius_m)
  movel([0.590936, -1.317764, -2.612347, -0.782278, 1.570796, 2.161732],accel_mss,speed_ms,0,blend_radius_m)
  movel([0.587426, -1.319203, -2.611455, -0.781732, 1.570796, 2.158222],accel_mss,speed_ms,0,blend_radius_m)
  movel([0.583959, -1.320247, -2.610806, -0.781337, 1.570796, 2.154755],accel_mss,speed_ms,0,blend_radius_m)
  movel([0.580533, -1.320927, -2.610382, -0.781080, 1.570796, 2.151330],accel_mss,speed_ms,0,blend_radius_m)
  movel([0.577159, -1.321270, -2.610168, -0.780951, 1.570796, 2.147955],accel_mss,speed_ms,0,blend_radius_m)
  movel([0.573835, -1.321303, -2.610148, -0.780939, 1.570796, 2.144632],accel_mss,speed_ms,0,blend_radius_m)
  movel([0.567369, -1.320535, -2.610626, -0.781228, 1.570796, 2.138165],accel_mss,speed_ms,0,blend_radius_m)
  movel([0.561177, -1.318829, -2.611687, -0.781873, 1.570796, 2.131974],accel_mss,speed_ms,0,blend_radius_m)
  movel([0.555312, -1.316374, -2.613207, -0.782809, 1.570796, 2.126108],accel_mss,speed_ms,0,blend_radius_m)
  movel([0.550235, -1.313463, -2.614998, -0.783928, 1.570796, 2.121031],accel_mss,speed_ms,0,blend_radius_m)
  movel([0.543806, -1.309606, -2.617354, -0.785428, 1.570796, 2.114603],accel_mss,speed_ms,0,blend_radius_m)
  movel([0.536275, -1.305789, -2.619667, -0.786933, 1.570796, 2.107071],accel_mss,speed_ms,0,blend_radius_m)
  movel([0.532183, -1.304205, -2.620622, -0.787562, 1.570796, 2.102979],accel_mss,speed_ms,0,blend_radius_m)
  movel([0.527925, -1.303003, -2.621344, -0.788043, 1.570796, 2.098721],accel_mss,speed_ms,0,blend_radius_m)
  movel([0.523547, -1.302302, -2.621764, -0.788323, 1.570796, 2.094343],accel_mss,speed_ms,0,blend_radius_m)
  movel([0.519094, -1.302222, -2.621811, -0.788355, 1.570796, 2.089890],accel_mss,speed_ms,0,blend_radius_m)
  movel([0.514617, -1.302881, -2.621417, -0.788091, 1.570796, 2.085413],accel_mss,speed_ms,0,blend_radius_m)
  movel([0.510166, -1.304387, -2.620512, -0.787490, 1.570796, 2.080963],accel_mss,speed_ms,0,blend_radius_m)
  movel([0.507970, -1.305492, -2.619847, -0.787050, 1.570796, 2.078766],accel_mss,speed_ms,0,blend_radius_m)
  movel([0.505801, -1.306846, -2.619029, -0.786514, 1.570796, 2.076598],accel_mss,speed_ms,0,blend_radius_m)
  movel([0.503666, -1.308465, -2.618048, -0.785876, 1.570796, 2.074463],accel_mss,speed_ms,0,blend_radius_m)
  movel([0.501574, -1.310360, -2.616896, -0.785134, 1.570796, 2.072371],accel_mss,speed_ms,0,blend_radius_m)
  movel([0.499533, -1.312540, -2.615563, -0.784285, 1.570796, 2.070329],accel_mss,speed_ms,0,blend_radius_m)
  movel([0.497547, -1.315019, -2.614042, -0.783328, 1.570796, 2.068344],accel_mss,speed_ms,0,blend_radius_m)
  movel([0.493776, -1.320905, -2.610396, -0.781088, 1.570796, 2.064572],accel_mss,speed_ms,0,blend_radius_m)
  movel([0.492676, -1.323790, -2.608592, -0.780007, 1.570796, 2.063472],accel_mss,speed_ms,0,blend_radius_m)
  movel([0.492116, -1.326662, -2.606785, -0.778942, 1.570796, 2.062912],accel_mss,speed_ms,0,blend_radius_m)
  movel([0.492132, -1.329496, -2.604991, -0.777902, 1.570796, 2.062928],accel_mss,speed_ms,0,blend_radius_m)
  movel([0.492763, -1.332260, -2.603231, -0.776898, 1.570796, 2.063560],accel_mss,speed_ms,0,blend_radius_m)
  movel([0.495919, -1.328700, -2.605496, -0.778193, 1.570796, 2.066715],accel_mss,speed_ms,0,blend_radius_m)
  movel([0.499273, -1.325443, -2.607553, -0.779393, 1.570796, 2.070069],accel_mss,speed_ms,0,blend_radius_m)
  movel([0.502788, -1.322505, -2.609397, -0.780488, 1.570796, 2.073584],accel_mss,speed_ms,0,blend_radius_m)
  movel([0.506430, -1.319903, -2.611020, -0.781467, 1.570796, 2.077227],accel_mss,speed_ms,0,blend_radius_m)
  movel([0.510162, -1.317651, -2.612417, -0.782321, 1.570796, 2.080959],accel_mss,speed_ms,0,blend_radius_m)
  movel([0.513944, -1.315764, -2.613583, -0.783042, 1.570796, 2.084740],accel_mss,speed_ms,0,blend_radius_m)
  movel([0.517738, -1.314254, -2.614513, -0.783623, 1.570796, 2.088534],accel_mss,speed_ms,0,blend_radius_m)
  movel([0.521504, -1.313136, -2.615199, -0.784054, 1.570796, 2.092301],accel_mss,speed_ms,0,blend_radius_m)
  movel([0.525206, -1.312420, -2.615637, -0.784332, 1.570796, 2.096002],accel_mss,speed_ms,0,blend_radius_m)
  movel([0.528805, -1.312117, -2.615822, -0.784449, 1.570796, 2.099601],accel_mss,speed_ms,0,blend_radius_m)
  movel([0.532262, -1.312238, -2.615749, -0.784402, 1.570796, 2.103058],accel_mss,speed_ms,0,blend_radius_m)
  movel([0.535540, -1.312789, -2.615411, -0.784189, 1.570796, 2.106336],accel_mss,speed_ms,0,blend_radius_m)
  movel([0.538599, -1.313780, -2.614803, -0.783806, 1.570796, 2.109396],accel_mss,speed_ms,0,blend_radius_m)
  movel([0.541405, -1.315212, -2.613923, -0.783254, 1.570796, 2.112202],accel_mss,speed_ms,0,blend_radius_m)
  movel([0.543925, -1.317092, -2.612763, -0.782534, 1.570796, 2.114722],accel_mss,speed_ms,0,blend_radius_m)
  movel([0.546119, -1.319421, -2.611319, -0.781649, 1.570796, 2.116915],accel_mss,speed_ms,0,blend_radius_m)
  movel([0.547610, -1.321618, -2.609951, -0.780820, 1.570796, 2.118406],accel_mss,speed_ms,0,blend_radius_m)
  movel([0.548743, -1.323966, -2.608481, -0.779942, 1.570796, 2.119539],accel_mss,speed_ms,0,blend_radius_m)
  movel([0.549534, -1.326441, -2.606924, -0.779024, 1.570796, 2.120330],accel_mss,speed_ms,0,blend_radius_m)
  movel([0.550003, -1.329021, -2.605292, -0.778076, 1.570796, 2.120799],accel_mss,speed_ms,0,blend_radius_m)
  movel([0.550035, -1.334417, -2.601850, -0.776122, 1.570796, 2.120831],accel_mss,speed_ms,0,blend_radius_m)
  movel([0.548981, -1.339990, -2.598253, -0.774145, 1.570796, 2.119777],accel_mss,speed_ms,0,blend_radius_m)
  movel([0.546971, -1.345591, -2.594596, -0.772202, 1.570796, 2.117767],accel_mss,speed_ms,0,blend_radius_m)
  movel([0.544134, -1.351073, -2.590975, -0.770341, 1.570796, 2.114930],accel_mss,speed_ms,0,blend_radius_m)
  movel([0.540590, -1.356299, -2.587484, -0.768607, 1.570796, 2.111387],accel_mss,speed_ms,0,blend_radius_m)
  movel([0.536457, -1.361143, -2.584214, -0.767033, 1.570796, 2.107253],accel_mss,speed_ms,0,blend_radius_m)
  movel([0.531843, -1.365476, -2.581261, -0.765652, 1.570796, 2.102640],accel_mss,speed_ms,0,blend_radius_m)
  movel([0.526854, -1.369175, -2.578719, -0.764495, 1.570796, 2.097650],accel_mss,speed_ms,0,blend_radius_m)
  movel([0.521584, -1.372126, -2.576677, -0.763586, 1.570796, 2.092380],accel_mss,speed_ms,0,blend_radius_m)
  movel([0.518875, -1.373280, -2.575875, -0.763234, 1.570796, 2.089671],accel_mss,speed_ms,0,blend_radius_m)
  movel([0.516127, -1.374205, -2.575231, -0.762953, 1.570796, 2.086923],accel_mss,speed_ms,0,blend_radius_m)
  movel([0.513357, -1.374881, -2.574760, -0.762748, 1.570796, 2.084153],accel_mss,speed_ms,0,blend_radius_m)
  movel([0.510571, -1.375294, -2.574472, -0.762624, 1.570796, 2.081367],accel_mss,speed_ms,0,blend_radius_m)
  movel([0.507780, -1.375426, -2.574379, -0.762584, 1.570796, 2.078576],accel_mss,speed_ms,0,blend_radius_m)
  movel([0.504993, -1.375267, -2.574490, -0.762632, 1.570796, 2.075790],accel_mss,speed_ms,0,blend_radius_m)
  movel([0.502225, -1.374795, -2.574820, -0.762774, 1.570796, 2.073021],accel_mss,speed_ms,0,blend_radius_m)
  movel([0.499481, -1.373996, -2.575377, -0.763016, 1.570796, 2.070277],accel_mss,speed_ms,0,blend_radius_m)
  movel([0.496772, -1.372853, -2.576172, -0.763364, 1.570796, 2.067569],accel_mss,speed_ms,0,blend_radius_m)
  movel([0.494108, -1.371345, -2.577218, -0.763825, 1.570796, 2.064904],accel_mss,speed_ms,0,blend_radius_m)
  movel([0.492284, -1.369743, -2.578327, -0.764319, 1.570796, 2.063081],accel_mss,speed_ms,0,blend_radius_m)
  movel([0.487818, -1.364744, -2.581761, -0.765884, 1.570796, 2.058614],accel_mss,speed_ms,0,blend_radius_m)
  movel([0.485054, -1.360877, -2.584394, -0.767118, 1.570796, 2.055850],accel_mss,speed_ms,0,blend_radius_m)
  movel([0.482180, -1.356035, -2.587661, -0.768693, 1.570796, 2.052977],accel_mss,speed_ms,0,blend_radius_m)
  movel([0.479388, -1.350163, -2.591578, -0.770647, 1.570796, 2.050184],accel_mss,speed_ms,0,blend_radius_m)
  movel([0.476871, -1.343196, -2.596165, -0.773028, 1.570796, 2.047667],accel_mss,speed_ms,0,blend_radius_m)
  movel([0.475594, -1.337993, -2.599547, -0.774849, 1.570796, 2.046390],accel_mss,speed_ms,0,blend_radius_m)
  movel([0.474967, -1.332973, -2.602775, -0.776641, 1.570796, 2.045764],accel_mss,speed_ms,0,blend_radius_m)
  movel([0.474919, -1.328153, -2.605842, -0.778394, 1.570796, 2.045716],accel_mss,speed_ms,0,blend_radius_m)
  movel([0.475384, -1.323549, -2.608743, -0.780097, 1.570796, 2.046180],accel_mss,speed_ms,0,blend_radius_m)
  movel([0.476283, -1.319183, -2.611467, -0.781739, 1.570796, 2.047079],accel_mss,speed_ms,0,blend_radius_m)
  movel([0.477540, -1.315076, -2.614007, -0.783306, 1.570796, 2.048336],accel_mss,speed_ms,0,blend_radius_m)
  movel([0.479079, -1.311252, -2.616351, -0.784786, 1.570796, 2.049876],accel_mss,speed_ms,0,blend_radius_m)
  movel([0.480818, -1.307731, -2.618493, -0.786165, 1.570796, 2.051615],accel_mss,speed_ms,0,blend_radius_m)
  movel([0.484560, -1.301701, -2.622123, -0.788564, 1.570796, 2.055356],accel_mss,speed_ms,0,blend_radius_m)
  movel([0.488091, -1.297174, -2.624818, -0.790397, 1.570796, 2.058887],accel_mss,speed_ms,0,blend_radius_m)
  movel([0.490715, -1.294336, -2.626494, -0.791559, 1.570796, 2.061511],accel_mss,speed_ms,0,blend_radius_m)
